// ---- SelfTests/TestCases/TestSuite_Preparation/Helper/PreparationResource.TcPOU
{region 'Documentation'}
(*!
<summary>Controlled local resource for Preparation selftests; only its FB call advances feedback. RequestValue records every command write, including repeated values. Initialize establishes a fresh fixture.</summary>
*)
{endregion}
FUNCTION_BLOCK PreparationResource
VAR_INPUT
    Available : BOOL := TRUE; //! Availability accepted on the next resource-body call.
    Fault : BOOL := FALSE; //! Technical fault accepted on the next resource-body call.
    Advance : BOOL := TRUE; //! FALSE holds feedback without cancelling the accepted request.
END_VAR
VAR
    FActualValue : DINT;
    FRequestedValue : DINT;
    FCommandWriteCount : UDINT;
    FAvailable : BOOL := TRUE;
    FFault : BOOL;
END_VAR

FAvailable := Available;
FFault := Fault;
IF NOT IsReady OR NOT Advance THEN
    RETURN;
END_IF;

IF FActualValue < FRequestedValue THEN
    FActualValue := FActualValue + 1;
ELSIF FActualValue > FRequestedValue THEN
    FActualValue := FActualValue - 1;
END_IF;

{region 'Documentation'}
(*!
<summary>Feedback after the last resource call.</summary>
*)
{endregion}
{attribute 'monitoring' := 'call'}
PROPERTY PUBLIC ActualValue : DINT //! Feedback after the last resource call.
GET // PUBLIC
ActualValue := FActualValue;
END_GET
END_PROPERTY

{region 'Documentation'}
(*!
<summary>Every RequestValue call since fixture initialization, including same-value writes.</summary>
*)
{endregion}
{attribute 'monitoring' := 'call'}
PROPERTY PUBLIC CommandWriteCount : UDINT //! Every RequestValue call since fixture initialization, including same-value writes.
GET // PUBLIC
CommandWriteCount := FCommandWriteCount;
END_GET
END_PROPERTY

{region 'Documentation'}
(*!
<summary>Fault accepted at the last resource call.</summary>
*)
{endregion}
{attribute 'monitoring' := 'call'}
PROPERTY PUBLIC HasError : BOOL //! Fault accepted at the last resource call.
GET // PUBLIC
HasError := FFault;
END_GET
END_PROPERTY

{region 'Documentation'}
(*!
<summary>Restores feedback and request together; fixture setup is not counted as a resource command.</summary>
*)
{endregion}
METHOD PUBLIC Initialize
VAR_INPUT
    InitialValue : DINT; //! Initial feedback and requested target; fixture initialization clears command-write evidence.
END_VAR
FActualValue := InitialValue;
FRequestedValue := InitialValue;
FCommandWriteCount := 0;
FAvailable := TRUE;
FFault := FALSE;
END_METHOD

{region 'Documentation'}
(*!
<summary>Current resource condition permits movement; independent of the target value.</summary>
*)
{endregion}
{attribute 'monitoring' := 'call'}
PROPERTY PUBLIC IsReady : BOOL //! Current resource condition permits movement; independent of the target value.
GET // PUBLIC
IsReady := FAvailable AND NOT FFault;
END_GET
END_PROPERTY

{region 'Documentation'}
(*!
<summary>Last requested target; accepting a command does not establish feedback.</summary>
*)
{endregion}
{attribute 'monitoring' := 'call'}
PROPERTY PUBLIC RequestedValue : DINT //! Last requested target; accepting a command does not establish feedback.
GET // PUBLIC
RequestedValue := FRequestedValue;
END_GET
END_PROPERTY

{region 'Documentation'}
(*!
<summary>Records one command write without changing feedback; a later advancing resource call processes it.</summary>
*)
{endregion}
METHOD PUBLIC RequestValue
VAR_INPUT
    Value : DINT; //! New requested target; this call records a command write without advancing feedback.
END_VAR
FRequestedValue := Value;
FCommandWriteCount := FCommandWriteCount + 1;
END_METHOD

END_FUNCTION_BLOCK

// ---- Framework/Assertions/POU/BasicTypes/DInt/AssertEqual_DInt.TcPOU
{region 'Documentation'}
(*!
<summary>Checks equality with the expected DINT value.</summary>
*)
{endregion}
FUNCTION_BLOCK AssertEqual_DInt EXTENDS AssertionBase
VAR_INPUT
    IN : DINT; //! Actual value checked or observed by this Assertion.
    Expected : DINT; //! Reference value for comparison with IN.
END_VAR

SUPER^();

{region 'Documentation'}
(*!
<summary>Check equality with the expected DINT value.</summary>
*)
{endregion}
METHOD PROTECTED Assert
VAR
    Message : STRING(GVL_Constants.MessageLength);
    ExpectedText : STRING(GVL_Constants.AssertionValueLength);
    ActualText : STRING(GVL_Constants.AssertionValueLength);
END_VAR
IF NOT EvaluationActive THEN
    RETURN;
END_IF;

IF Result = E_Result.Error THEN
    RETURN;
END_IF;

IF Result = E_Result.Failed THEN
    RETURN;
END_IF;

IF IN <> Expected THEN
    ExpectedText := DINT_TO_STRING(Expected);
    ActualText := DINT_TO_STRING(IN);
    Message := CONCAT('Assertion failed: values are not equal. Expected = ',
        ExpectedText);
    Message := CONCAT(Message, ', Actual = ');
    Message := CONCAT(Message, ActualText);
    Message := CONCAT(Message, '.');
    Fail(Message := Message);
    RETURN;
END_IF;

Pass();
END_METHOD

END_FUNCTION_BLOCK

// ---- SelfTests/TestCases/TestSuite_Preparation/Test_PreparationReachesTarget.TcPOU
{region 'Documentation'}
(*!
<summary>Checks real request/feedback separation, multi-cycle target acquisition and already-reached behavior.</summary>
*)
{endregion}
FUNCTION_BLOCK Test_PreparationReachesTarget EXTENDS TestCaseBase
VAR
    FSubject : Prepare_ValueAtTarget;
    FResource : PreparationResource;
    FView : I_Preparation;
    FAlreadyAtTarget : Prepare_ValueAtTarget;
    FObserved : ST_PreparationStatus;
    FExpected : ST_PreparationStatus;
    FObservedEnabled : BOOL;
    FExpectedEnabled : BOOL;
    FCheckPerformed : BOOL;
    FObservedCommandWrites : UDINT;
    FExpectedCommandWrites : UDINT;
    FObservedActualValue : DINT;
    FExpectedActualValue : DINT;
    FObservedRequestedValue : DINT;
    FExpectedRequestedValue : DINT;
    FCheckDiagnosticState : AssertEqual_Int;
    FCheckExecutionStatus : AssertEqual_Int;
    FCheckReady : AssertEqual_Bool;
    FCheckRunning : AssertEqual_Bool;
    FCheckCompleted : AssertEqual_Bool;
    FCheckError : AssertEqual_Bool;
    FCheckEnabled : AssertEqual_Bool;
    FCheckCommandWrites : AssertEqual_UDInt;
    FCheckActualValue : AssertEqual_DInt;
    FCheckRequestedValue : AssertEqual_DInt;
END_VAR
VAR CONSTANT
    CommandAccepted : E_State := E_State.Running;
    ProgressObserved : E_State := E_State.Running + 1;
    TargetReached : E_State := E_State.Running + 2;
    RepeatedCompletion : E_State := E_State.Running + 3;
    AlreadyAtTarget : E_State := E_State.Running + 4;
END_VAR

SUPER^();

{region 'Documentation'}
(*!
<summary>Contributes all owned Assertion results without executing the subjects.</summary>
*)
{endregion}
METHOD PROTECTED AggregateResults
VAR_INPUT
    Aggregator : I_ResultAggregator; //! Borrowed result sink owned by the outer Test Case; add this test's checking Assertions without resetting or retaining the sink.
END_VAR
Aggregator.AddProvider(Provider := FCheckDiagnosticState);
Aggregator.AddProvider(Provider := FCheckExecutionStatus);
Aggregator.AddProvider(Provider := FCheckReady);
Aggregator.AddProvider(Provider := FCheckRunning);
Aggregator.AddProvider(Provider := FCheckCompleted);
Aggregator.AddProvider(Provider := FCheckError);
Aggregator.AddProvider(Provider := FCheckEnabled);
Aggregator.AddProvider(Provider := FCheckCommandWrites);
Aggregator.AddProvider(Provider := FCheckActualValue);
Aggregator.AddProvider(Provider := FCheckRequestedValue);
END_METHOD

{region 'Documentation'}
(*!
<summary>Requires valid base configuration and every owned Assertion.</summary>
*)
{endregion}
METHOD PROTECTED CheckInitialization : BOOL //! TRUE when the inherited initialization check and this concrete fixture check both accept the setup.
CheckInitialization := FALSE;
IF NOT SUPER^.CheckInitialization() THEN
    RETURN;
END_IF;
IF NOT FCheckDiagnosticState.IsInitialized
    OR NOT FCheckExecutionStatus.IsInitialized
    OR NOT FCheckReady.IsInitialized
    OR NOT FCheckRunning.IsInitialized
    OR NOT FCheckCompleted.IsInitialized
    OR NOT FCheckError.IsInitialized
    OR NOT FCheckEnabled.IsInitialized
    OR NOT FCheckCommandWrites.IsInitialized
    OR NOT FCheckActualValue.IsInitialized
    OR NOT FCheckRequestedValue.IsInitialized THEN
    RETURN;
END_IF;

CheckInitialization := TRUE;
END_METHOD

{region 'Documentation'}
(*!
<summary>Configures this scenario, its local subjects and named Assertions.</summary>
*)
{endregion}
METHOD PROTECTED Configure
FPreparationStateCount := 0;
FTestStateCount := 5;
FCheckPerformed := FALSE;
FResource.Initialize(InitialValue := 2);
FSubject.Initialize(Resource := FResource);
FAlreadyAtTarget.Initialize(Resource := FResource);
FView := FSubject;

FCheckDiagnosticState.Initialize(Parent := THIS^,
    AssertionName := 'DiagnosticState');
FCheckExecutionStatus.Initialize(Parent := THIS^,
    AssertionName := 'ExecutionStatus');
FCheckReady.Initialize(Parent := THIS^,
    AssertionName := 'Ready');
FCheckRunning.Initialize(Parent := THIS^,
    AssertionName := 'Running');
FCheckCompleted.Initialize(Parent := THIS^,
    AssertionName := 'Completed');
FCheckError.Initialize(Parent := THIS^,
    AssertionName := 'Error');
FCheckEnabled.Initialize(Parent := THIS^,
    AssertionName := 'Enabled');
FCheckCommandWrites.Initialize(Parent := THIS^,
    AssertionName := 'CommandWrites');
FCheckActualValue.Initialize(Parent := THIS^,
    AssertionName := 'ActualValue');
FCheckRequestedValue.Initialize(Parent := THIS^,
    AssertionName := 'RequestedValue');
END_METHOD

{region 'Documentation'}
(*!
<summary>Ends scenario processing without issuing further resource commands.</summary>
*)
{endregion}
METHOD PROTECTED ProcessAbort
VAR_INPUT
    Enable : BOOL; //! Phase permission supplied by the owning Test Case; FALSE does not authorize progression, while observation may continue.
END_VAR
IF Enable THEN
    CompleteAbort();
END_IF;
END_METHOD

{region 'Documentation'}
(*!
<summary>Compares independent expected values with the captured observations; called when disabled as well.</summary>
*)
{endregion}
METHOD PROTECTED ProcessAssertions
VAR_INPUT
    Enable : BOOL; //! Phase permission supplied by the owning Test Case; FALSE does not authorize progression, while observation may continue.
END_VAR
FCheckDiagnosticState(Enable := Enable,
    State := State,
    IN := TO_INT(FObserved.State),
    Expected := TO_INT(FExpected.State));

FCheckExecutionStatus(Enable := Enable,
    State := State,
    IN := TO_INT(FObserved.ExecutionStatus),
    Expected := TO_INT(FExpected.ExecutionStatus));

FCheckReady(Enable := Enable,
    State := State,
    IN := FObserved.Ready,
    Expected := FExpected.Ready);

FCheckRunning(Enable := Enable,
    State := State,
    IN := FObserved.Running,
    Expected := FExpected.Running);

FCheckCompleted(Enable := Enable,
    State := State,
    IN := FObserved.Completed,
    Expected := FExpected.Completed);

FCheckError(Enable := Enable,
    State := State,
    IN := FObserved.Error,
    Expected := FExpected.Error);

FCheckEnabled(Enable := Enable,
    State := State,
    IN := FObservedEnabled,
    Expected := FExpectedEnabled);

FCheckCommandWrites(Enable := Enable,
    State := State,
    IN := FObservedCommandWrites,
    Expected := FExpectedCommandWrites);

FCheckActualValue(Enable := Enable,
    State := State,
    IN := FObservedActualValue,
    Expected := FExpectedActualValue);

FCheckRequestedValue(Enable := Enable,
    State := State,
    IN := FObservedRequestedValue,
    Expected := FExpectedRequestedValue);

IF Enable
    AND FCheckDiagnosticState.EvaluationActive
    AND FCheckExecutionStatus.EvaluationActive
    AND FCheckReady.EvaluationActive
    AND FCheckRunning.EvaluationActive
    AND FCheckCompleted.EvaluationActive
    AND FCheckError.EvaluationActive
    AND FCheckEnabled.EvaluationActive
    AND FCheckCommandWrites.EvaluationActive
    AND FCheckActualValue.EvaluationActive
    AND FCheckRequestedValue.EvaluationActive THEN
    FCheckPerformed := TRUE;
END_IF;
END_METHOD

{region 'Documentation'}
(*!
<summary>Subjects are exercised by the test, not used as its start prerequisite.</summary>
*)
{endregion}
METHOD PROTECTED ProcessPreparations
VAR_INPUT
    // SA0033: Required hook; this scenario has no Preparation phase.
    {attribute 'analysis' := '-33'}
    Enable : BOOL; //! Phase permission supplied by the owning Test Case; FALSE does not authorize progression, while observation may continue.
END_VAR
END_METHOD

{region 'Documentation'}
(*!
<summary>Restores repeatable fixture state and resets Assertions before returning to Idle.</summary>
*)
{endregion}
METHOD PROTECTED ProcessReset
FCheckPerformed := FALSE;
FResource.Initialize(InitialValue := 2);
FSubject.Initialize(Resource := FResource);
FAlreadyAtTarget.Initialize(Resource := FResource);
FView := FSubject;
FCheckDiagnosticState.Reset();
FCheckExecutionStatus.Reset();
FCheckReady.Reset();
FCheckRunning.Reset();
FCheckCompleted.Reset();
FCheckError.Reset();
FCheckEnabled.Reset();
FCheckCommandWrites.Reset();
FCheckActualValue.Reset();
FCheckRequestedValue.Reset();
CompleteReset();
END_METHOD

{region 'Documentation'}
(*!
<summary>Exercises one named scenario step per call; advances only after actual Assertion evaluation.</summary>
*)
{endregion}
METHOD PROTECTED ProcessTests
VAR_INPUT
    Enable : BOOL; //! Phase permission supplied by the owning Test Case; FALSE does not authorize progression, while observation may continue.
END_VAR
IF NOT Enable THEN
    RETURN;
END_IF;

IF FCheckPerformed THEN
    FCheckPerformed := FALSE;
    IF State = AlreadyAtTarget THEN
        CompleteTests();
        RETURN;
    END_IF;
    NextTestState();
    IF NOT IsTestingActive THEN
        RETURN;
    END_IF;
END_IF;

CASE State OF
    CommandAccepted:
        FResource(Available := TRUE,
            Fault := FALSE,
            Advance := FALSE);
        FSubject(Enable := TRUE,
            TargetValue := 0);
        FExpected.State := E_State.Running;
        FExpected.ExecutionStatus := E_ExecutionStatus.Running;
        FExpected.Ready := FALSE;
        FExpected.Running := TRUE;
        FExpected.Completed := FALSE;
        FExpected.Error := FALSE;
        FExpectedEnabled := TRUE;
        FExpectedCommandWrites := 1;
        FExpectedActualValue := 2;
        FExpectedRequestedValue := 0;

    ProgressObserved:
        FResource(Available := TRUE,
            Fault := FALSE,
            Advance := TRUE);
        FSubject(Enable := TRUE,
            TargetValue := 0);
        FExpected.State := E_State.Running;
        FExpected.ExecutionStatus := E_ExecutionStatus.Running;
        FExpected.Ready := FALSE;
        FExpected.Running := TRUE;
        FExpected.Completed := FALSE;
        FExpected.Error := FALSE;
        FExpectedEnabled := TRUE;
        FExpectedCommandWrites := 1;
        FExpectedActualValue := 1;
        FExpectedRequestedValue := 0;

    TargetReached:
        FResource(Available := TRUE,
            Fault := FALSE,
            Advance := TRUE);
        FSubject(Enable := TRUE,
            TargetValue := 0);
        FExpected.State := E_State.Completed;
        FExpected.ExecutionStatus := E_ExecutionStatus.Completed;
        FExpected.Ready := TRUE;
        FExpected.Running := FALSE;
        FExpected.Completed := TRUE;
        FExpected.Error := FALSE;
        FExpectedEnabled := TRUE;
        FExpectedCommandWrites := 1;
        FExpectedActualValue := 0;
        FExpectedRequestedValue := 0;

    RepeatedCompletion:
        FResource(Available := TRUE,
            Fault := FALSE,
            Advance := TRUE);
        FSubject(Enable := TRUE,
            TargetValue := 0);
        FExpected.State := E_State.Completed;
        FExpected.ExecutionStatus := E_ExecutionStatus.Completed;
        FExpected.Ready := TRUE;
        FExpected.Running := FALSE;
        FExpected.Completed := TRUE;
        FExpected.Error := FALSE;
        FExpectedEnabled := TRUE;
        FExpectedCommandWrites := 1;
        FExpectedActualValue := 0;
        FExpectedRequestedValue := 0;

    AlreadyAtTarget:
        FResource(Available := TRUE,
            Fault := FALSE,
            Advance := TRUE);
        FAlreadyAtTarget(Enable := TRUE,
            TargetValue := 0);
        FView := FAlreadyAtTarget;
        FExpected.State := E_State.Completed;
        FExpected.ExecutionStatus := E_ExecutionStatus.Completed;
        FExpected.Ready := TRUE;
        FExpected.Running := FALSE;
        FExpected.Completed := TRUE;
        FExpected.Error := FALSE;
        FExpectedEnabled := TRUE;
        FExpectedCommandWrites := 1;
        FExpectedActualValue := 0;
        FExpectedRequestedValue := 0;

ELSE
    Error(Message := 'Unexpected Preparation test state.');
    RETURN;
END_CASE;

FObserved := FView.Status;
IF State = AlreadyAtTarget THEN
    FObservedEnabled := FAlreadyAtTarget.Enabled;
ELSE
    FObservedEnabled := FSubject.Enabled;
END_IF;

FObservedCommandWrites := FResource.CommandWriteCount;
FObservedActualValue := FResource.ActualValue;
FObservedRequestedValue := FResource.RequestedValue;
END_METHOD

END_FUNCTION_BLOCK

// ---- SelfTests/TestCases/TestSuite_Preparation/Test_PreparationDisableAndReenable.TcPOU
{region 'Documentation'}
(*!
<summary>Checks that disabling discards local stage progress without cancelling the accepted resource command.</summary>
*)
{endregion}
FUNCTION_BLOCK Test_PreparationDisableAndReenable EXTENDS TestCaseBase
VAR
    FSubject : Prepare_ZeroViaOne;
    FResource : PreparationResource;
    FView : I_Preparation;
    FObserved : ST_PreparationStatus;
    FExpected : ST_PreparationStatus;
    FObservedEnabled : BOOL;
    FExpectedEnabled : BOOL;
    FCheckPerformed : BOOL;
    FObservedCommandWrites : UDINT;
    FExpectedCommandWrites : UDINT;
    FObservedActualValue : DINT;
    FExpectedActualValue : DINT;
    FObservedRequestedValue : DINT;
    FExpectedRequestedValue : DINT;
    FCheckDiagnosticState : AssertEqual_Int;
    FCheckExecutionStatus : AssertEqual_Int;
    FCheckReady : AssertEqual_Bool;
    FCheckRunning : AssertEqual_Bool;
    FCheckCompleted : AssertEqual_Bool;
    FCheckError : AssertEqual_Bool;
    FCheckEnabled : AssertEqual_Bool;
    FCheckCommandWrites : AssertEqual_UDInt;
    FCheckActualValue : AssertEqual_DInt;
    FCheckRequestedValue : AssertEqual_DInt;
END_VAR
VAR CONSTANT
    IntermediateRequested : E_State := E_State.Running;
    DisableDuringMovement : E_State := E_State.Running + 1;
    AcceptedRequestContinues : E_State := E_State.Running + 2;
    ResourceChangedWhileDisabled : E_State := E_State.Running + 3;
    ReenableFromCurrentFeedback : E_State := E_State.Running + 4;
    IntermediateApproached : E_State := E_State.Running + 5;
    FinalTargetRequested : E_State := E_State.Running + 6;
    FinalTargetReached : E_State := E_State.Running + 7;
END_VAR

SUPER^();

{region 'Documentation'}
(*!
<summary>Contributes all owned Assertion results without executing the subjects.</summary>
*)
{endregion}
METHOD PROTECTED AggregateResults
VAR_INPUT
    Aggregator : I_ResultAggregator; //! Borrowed result sink owned by the outer Test Case; add this test's checking Assertions without resetting or retaining the sink.
END_VAR
Aggregator.AddProvider(Provider := FCheckDiagnosticState);
Aggregator.AddProvider(Provider := FCheckExecutionStatus);
Aggregator.AddProvider(Provider := FCheckReady);
Aggregator.AddProvider(Provider := FCheckRunning);
Aggregator.AddProvider(Provider := FCheckCompleted);
Aggregator.AddProvider(Provider := FCheckError);
Aggregator.AddProvider(Provider := FCheckEnabled);
Aggregator.AddProvider(Provider := FCheckCommandWrites);
Aggregator.AddProvider(Provider := FCheckActualValue);
Aggregator.AddProvider(Provider := FCheckRequestedValue);
END_METHOD

{region 'Documentation'}
(*!
<summary>Requires valid base configuration and every owned Assertion.</summary>
*)
{endregion}
METHOD PROTECTED CheckInitialization : BOOL //! TRUE when the inherited initialization check and this concrete fixture check both accept the setup.
CheckInitialization := FALSE;
IF NOT SUPER^.CheckInitialization() THEN
    RETURN;
END_IF;
IF NOT FCheckDiagnosticState.IsInitialized
    OR NOT FCheckExecutionStatus.IsInitialized
    OR NOT FCheckReady.IsInitialized
    OR NOT FCheckRunning.IsInitialized
    OR NOT FCheckCompleted.IsInitialized
    OR NOT FCheckError.IsInitialized
    OR NOT FCheckEnabled.IsInitialized
    OR NOT FCheckCommandWrites.IsInitialized
    OR NOT FCheckActualValue.IsInitialized
    OR NOT FCheckRequestedValue.IsInitialized THEN
    RETURN;
END_IF;

CheckInitialization := TRUE;
END_METHOD

{region 'Documentation'}
(*!
<summary>Configures this scenario, its local subjects and named Assertions.</summary>
*)
{endregion}
METHOD PROTECTED Configure
FPreparationStateCount := 0;
FTestStateCount := 8;
FCheckPerformed := FALSE;
FResource.Initialize(InitialValue := 3);
FSubject.Initialize(Resource := FResource);
FView := FSubject;

FCheckDiagnosticState.Initialize(Parent := THIS^,
    AssertionName := 'DiagnosticState');
FCheckExecutionStatus.Initialize(Parent := THIS^,
    AssertionName := 'ExecutionStatus');
FCheckReady.Initialize(Parent := THIS^,
    AssertionName := 'Ready');
FCheckRunning.Initialize(Parent := THIS^,
    AssertionName := 'Running');
FCheckCompleted.Initialize(Parent := THIS^,
    AssertionName := 'Completed');
FCheckError.Initialize(Parent := THIS^,
    AssertionName := 'Error');
FCheckEnabled.Initialize(Parent := THIS^,
    AssertionName := 'Enabled');
FCheckCommandWrites.Initialize(Parent := THIS^,
    AssertionName := 'CommandWrites');
FCheckActualValue.Initialize(Parent := THIS^,
    AssertionName := 'ActualValue');
FCheckRequestedValue.Initialize(Parent := THIS^,
    AssertionName := 'RequestedValue');
END_METHOD

{region 'Documentation'}
(*!
<summary>Ends scenario processing without issuing further resource commands.</summary>
*)
{endregion}
METHOD PROTECTED ProcessAbort
VAR_INPUT
    Enable : BOOL; //! Phase permission supplied by the owning Test Case; FALSE does not authorize progression, while observation may continue.
END_VAR
IF Enable THEN
    CompleteAbort();
END_IF;
END_METHOD

{region 'Documentation'}
(*!
<summary>Compares independent expected values with the captured observations; called when disabled as well.</summary>
*)
{endregion}
METHOD PROTECTED ProcessAssertions
VAR_INPUT
    Enable : BOOL; //! Phase permission supplied by the owning Test Case; FALSE does not authorize progression, while observation may continue.
END_VAR
FCheckDiagnosticState(Enable := Enable,
    State := State,
    IN := TO_INT(FObserved.State),
    Expected := TO_INT(FExpected.State));

FCheckExecutionStatus(Enable := Enable,
    State := State,
    IN := TO_INT(FObserved.ExecutionStatus),
    Expected := TO_INT(FExpected.ExecutionStatus));

FCheckReady(Enable := Enable,
    State := State,
    IN := FObserved.Ready,
    Expected := FExpected.Ready);

FCheckRunning(Enable := Enable,
    State := State,
    IN := FObserved.Running,
    Expected := FExpected.Running);

FCheckCompleted(Enable := Enable,
    State := State,
    IN := FObserved.Completed,
    Expected := FExpected.Completed);

FCheckError(Enable := Enable,
    State := State,
    IN := FObserved.Error,
    Expected := FExpected.Error);

FCheckEnabled(Enable := Enable,
    State := State,
    IN := FObservedEnabled,
    Expected := FExpectedEnabled);

FCheckCommandWrites(Enable := Enable,
    State := State,
    IN := FObservedCommandWrites,
    Expected := FExpectedCommandWrites);

FCheckActualValue(Enable := Enable,
    State := State,
    IN := FObservedActualValue,
    Expected := FExpectedActualValue);

FCheckRequestedValue(Enable := Enable,
    State := State,
    IN := FObservedRequestedValue,
    Expected := FExpectedRequestedValue);

IF Enable
    AND FCheckDiagnosticState.EvaluationActive
    AND FCheckExecutionStatus.EvaluationActive
    AND FCheckReady.EvaluationActive
    AND FCheckRunning.EvaluationActive
    AND FCheckCompleted.EvaluationActive
    AND FCheckError.EvaluationActive
    AND FCheckEnabled.EvaluationActive
    AND FCheckCommandWrites.EvaluationActive
    AND FCheckActualValue.EvaluationActive
    AND FCheckRequestedValue.EvaluationActive THEN
    FCheckPerformed := TRUE;
END_IF;
END_METHOD

{region 'Documentation'}
(*!
<summary>Subjects are exercised by the test, not used as its start prerequisite.</summary>
*)
{endregion}
METHOD PROTECTED ProcessPreparations
VAR_INPUT
    // SA0033: Required hook; this scenario has no Preparation phase.
    {attribute 'analysis' := '-33'}
    Enable : BOOL; //! Phase permission supplied by the owning Test Case; FALSE does not authorize progression, while observation may continue.
END_VAR
END_METHOD

{region 'Documentation'}
(*!
<summary>Restores repeatable fixture state and resets Assertions before returning to Idle.</summary>
*)
{endregion}
METHOD PROTECTED ProcessReset
FCheckPerformed := FALSE;
FResource.Initialize(InitialValue := 3);
FSubject.Initialize(Resource := FResource);
FView := FSubject;
FCheckDiagnosticState.Reset();
FCheckExecutionStatus.Reset();
FCheckReady.Reset();
FCheckRunning.Reset();
FCheckCompleted.Reset();
FCheckError.Reset();
FCheckEnabled.Reset();
FCheckCommandWrites.Reset();
FCheckActualValue.Reset();
FCheckRequestedValue.Reset();
CompleteReset();
END_METHOD

{region 'Documentation'}
(*!
<summary>Exercises one named scenario step per call; advances only after actual Assertion evaluation.</summary>
*)
{endregion}
METHOD PROTECTED ProcessTests
VAR_INPUT
    Enable : BOOL; //! Phase permission supplied by the owning Test Case; FALSE does not authorize progression, while observation may continue.
END_VAR
IF NOT Enable THEN
    RETURN;
END_IF;

IF FCheckPerformed THEN
    FCheckPerformed := FALSE;
    IF State = FinalTargetReached THEN
        CompleteTests();
        RETURN;
    END_IF;
    NextTestState();
    IF NOT IsTestingActive THEN
        RETURN;
    END_IF;
END_IF;

CASE State OF
    IntermediateRequested:
        FResource(Available := TRUE,
            Fault := FALSE,
            Advance := FALSE);
        FSubject(Enable := TRUE);
        FExpected.State := E_State.Preparing;
        FExpected.ExecutionStatus := E_ExecutionStatus.Running;
        FExpected.Ready := FALSE;
        FExpected.Running := TRUE;
        FExpected.Completed := FALSE;
        FExpected.Error := FALSE;
        FExpectedEnabled := TRUE;
        FExpectedCommandWrites := 1;
        FExpectedActualValue := 3;
        FExpectedRequestedValue := 1;

    DisableDuringMovement:
        FResource(Available := TRUE,
            Fault := FALSE,
            Advance := TRUE);
        FSubject(Enable := FALSE);
        FExpected.State := E_State.Idle;
        FExpected.ExecutionStatus := E_ExecutionStatus.Idle;
        FExpected.Ready := TRUE;
        FExpected.Running := FALSE;
        FExpected.Completed := FALSE;
        FExpected.Error := FALSE;
        FExpectedEnabled := FALSE;
        FExpectedCommandWrites := 1;
        FExpectedActualValue := 2;
        FExpectedRequestedValue := 1;

    AcceptedRequestContinues:
        FResource(Available := TRUE,
            Fault := FALSE,
            Advance := TRUE);
        FSubject(Enable := FALSE);
        FExpected.State := E_State.Idle;
        FExpected.ExecutionStatus := E_ExecutionStatus.Idle;
        FExpected.Ready := TRUE;
        FExpected.Running := FALSE;
        FExpected.Completed := FALSE;
        FExpected.Error := FALSE;
        FExpectedEnabled := FALSE;
        FExpectedCommandWrites := 1;
        FExpectedActualValue := 1;
        FExpectedRequestedValue := 1;

    ResourceChangedWhileDisabled:
        FResource.RequestValue(Value := 3);
        FResource(Available := TRUE,
            Fault := FALSE,
            Advance := TRUE);
        FSubject(Enable := FALSE);
        FExpected.State := E_State.Idle;
        FExpected.ExecutionStatus := E_ExecutionStatus.Idle;
        FExpected.Ready := TRUE;
        FExpected.Running := FALSE;
        FExpected.Completed := FALSE;
        FExpected.Error := FALSE;
        FExpectedEnabled := FALSE;
        FExpectedCommandWrites := 2;
        FExpectedActualValue := 2;
        FExpectedRequestedValue := 3;

    ReenableFromCurrentFeedback:
        FResource(Available := TRUE,
            Fault := FALSE,
            Advance := TRUE);
        FSubject(Enable := TRUE);
        FExpected.State := E_State.Preparing;
        FExpected.ExecutionStatus := E_ExecutionStatus.Running;
        FExpected.Ready := FALSE;
        FExpected.Running := TRUE;
        FExpected.Completed := FALSE;
        FExpected.Error := FALSE;
        FExpectedEnabled := TRUE;
        FExpectedCommandWrites := 3;
        FExpectedActualValue := 3;
        FExpectedRequestedValue := 1;

    IntermediateApproached:
        FResource(Available := TRUE,
            Fault := FALSE,
            Advance := TRUE);
        FSubject(Enable := TRUE);
        FExpected.State := E_State.Preparing;
        FExpected.ExecutionStatus := E_ExecutionStatus.Running;
        FExpected.Ready := FALSE;
        FExpected.Running := TRUE;
        FExpected.Completed := FALSE;
        FExpected.Error := FALSE;
        FExpectedEnabled := TRUE;
        FExpectedCommandWrites := 3;
        FExpectedActualValue := 2;
        FExpectedRequestedValue := 1;

    FinalTargetRequested:
        FResource(Available := TRUE,
            Fault := FALSE,
            Advance := TRUE);
        FSubject(Enable := TRUE);
        FExpected.State := E_State.Running;
        FExpected.ExecutionStatus := E_ExecutionStatus.Running;
        FExpected.Ready := FALSE;
        FExpected.Running := TRUE;
        FExpected.Completed := FALSE;
        FExpected.Error := FALSE;
        FExpectedEnabled := TRUE;
        FExpectedCommandWrites := 4;
        FExpectedActualValue := 1;
        FExpectedRequestedValue := 0;

    FinalTargetReached:
        FResource(Available := TRUE,
            Fault := FALSE,
            Advance := TRUE);
        FSubject(Enable := TRUE);
        FExpected.State := E_State.Completed;
        FExpected.ExecutionStatus := E_ExecutionStatus.Completed;
        FExpected.Ready := TRUE;
        FExpected.Running := FALSE;
        FExpected.Completed := TRUE;
        FExpected.Error := FALSE;
        FExpectedEnabled := TRUE;
        FExpectedCommandWrites := 4;
        FExpectedActualValue := 0;
        FExpectedRequestedValue := 0;

ELSE
    Error(Message := 'Unexpected Preparation test state.');
    RETURN;
END_CASE;

FObserved := FView.Status;
FObservedEnabled := FSubject.Enabled;

FObservedCommandWrites := FResource.CommandWriteCount;
FObservedActualValue := FResource.ActualValue;
FObservedRequestedValue := FResource.RequestedValue;
END_METHOD

END_FUNCTION_BLOCK

// ---- SelfTests/TestCases/TestSuite_Preparation/Helper/Prepare_ZeroViaOne.TcPOU
{region 'Documentation'}
(*!
<summary>Stateful local Preparation: establish value one before commanding zero. Disabled calls discard local progress without cancelling the resource request.</summary>
*)
{endregion}
FUNCTION_BLOCK Prepare_ZeroViaOne EXTENDS PreparationBase
VAR
    FResource : REFERENCE TO PreparationResource;
    FProgress : E_State := E_State.Idle;
END_VAR

VAR CONSTANT
    IntermediateValue : DINT := 1;
    TargetValue : DINT := 0;
END_VAR

SUPER^();

{region 'Documentation'}
(*!
<summary>Binds a static test-owned resource and clears local sequence progress.</summary>
*)
{endregion}
METHOD PUBLIC Initialize
VAR_IN_OUT
    // SA0167: Borrowed static resource, not a temporary instance.
    {attribute 'analysis' := '-167'}
    Resource : PreparationResource; //! Borrowed static resource retained by reference; keep it alive and stable for all preparation calls.
END_VAR
FResource REF= Resource;
FProgress := E_State.Idle;
END_METHOD

{region 'Documentation'}
(*!
<summary>Observes current feedback; enabling permits the two-stage resource sequence.</summary>
*)
{endregion}
METHOD PROTECTED Prepare
IF NOT Enabled THEN
    FProgress := E_State.Idle;
END_IF;
IF NOT __ISVALIDREF(FResource) THEN
    UpdateStatus(State := E_State.Error,
        ExecutionStatus := E_ExecutionStatus.Error,
        Ready := FALSE);
    RETURN;
END_IF;
IF FResource.HasError THEN
    UpdateStatus(State := E_State.Error,
        ExecutionStatus := E_ExecutionStatus.Error,
        Ready := FALSE);
    RETURN;
END_IF;

IF (FResource.ActualValue = TargetValue) AND (FResource.RequestedValue = TargetValue) THEN
    UpdateStatus(State := E_State.Completed,
        ExecutionStatus := E_ExecutionStatus.Completed,
        Ready := FResource.IsReady);
ELSIF Enabled AND FResource.IsReady THEN
    StateMachine();
    IF FProgress = E_State.Error THEN
        UpdateStatus(State := E_State.Error,
            ExecutionStatus := E_ExecutionStatus.Error,
            Ready := FALSE);
    ELSE
        UpdateStatus(State := FProgress,
            ExecutionStatus := E_ExecutionStatus.Running,
            Ready := FALSE);
    END_IF;
ELSIF FResource.IsReady THEN
    UpdateStatus(State := E_State.Idle,
        ExecutionStatus := E_ExecutionStatus.Idle,
        Ready := TRUE);
ELSE
    UpdateStatus(State := E_State.Idle,
        ExecutionStatus := E_ExecutionStatus.NotReady,
        Ready := FALSE);
END_IF;
END_METHOD

{region 'Documentation'}
(*!
<summary>Advances at most one resource stage per call; no feedback simulation.</summary>
*)
{endregion}
METHOD PRIVATE StateMachine
CASE FProgress OF
    E_State.Idle:
        IF FResource.ActualValue = IntermediateValue THEN
            FResource.RequestValue(Value := TargetValue);
            FProgress := E_State.Running;
        ELSE
            FResource.RequestValue(Value := IntermediateValue);
            FProgress := E_State.Preparing;
        END_IF;

    E_State.Preparing:
        IF FResource.ActualValue = IntermediateValue THEN
            FResource.RequestValue(Value := TargetValue);
            FProgress := E_State.Running;
        END_IF;

    E_State.Running:
        RETURN;
ELSE
    FProgress := E_State.Error;
END_CASE;
END_METHOD

END_FUNCTION_BLOCK

// ---- SelfTests/TestCases/TestSuite_Preparation/Test_PreparationCompletionTracksTarget.TcPOU
{region 'Documentation'}
(*!
<summary>Checks real Preparation-to-test handover; loss of Ready/Completed does not restart or block the active Test Case.</summary>
*)
{endregion}
FUNCTION_BLOCK Test_PreparationCompletionTracksTarget EXTENDS TestCaseBase
VAR
    FSubject : Prepare_ValueAtTarget;
    FResource : PreparationResource;
    FView : I_Preparation;
    FResourceAvailable : BOOL := TRUE;
    FObserved : ST_PreparationStatus;
    FExpected : ST_PreparationStatus;
    FObservedEnabled : BOOL;
    FExpectedEnabled : BOOL;
    FCheckPerformed : BOOL;
    FObservedCommandWrites : UDINT;
    FExpectedCommandWrites : UDINT;
    FObservedActualValue : DINT;
    FExpectedActualValue : DINT;
    FObservedRequestedValue : DINT;
    FExpectedRequestedValue : DINT;
    FCheckDiagnosticState : AssertEqual_Int;
    FCheckExecutionStatus : AssertEqual_Int;
    FCheckReady : AssertEqual_Bool;
    FCheckRunning : AssertEqual_Bool;
    FCheckCompleted : AssertEqual_Bool;
    FCheckError : AssertEqual_Bool;
    FCheckEnabled : AssertEqual_Bool;
    FCheckCommandWrites : AssertEqual_UDInt;
    FCheckActualValue : AssertEqual_DInt;
    FCheckRequestedValue : AssertEqual_DInt;
    FCheckTestingActive : AssertEqual_Bool;
END_VAR
VAR CONSTANT
    PreparationHandedOver : E_State := E_State.Running;
    TargetAndReadinessLost : E_State := E_State.Running + 1;
    TestingContinues : E_State := E_State.Running + 2;
END_VAR

SUPER^();

{region 'Documentation'}
(*!
<summary>Contributes all owned Assertion results without executing the subjects.</summary>
*)
{endregion}
METHOD PROTECTED AggregateResults
VAR_INPUT
    Aggregator : I_ResultAggregator; //! Borrowed result sink owned by the outer Test Case; add this test's checking Assertions without resetting or retaining the sink.
END_VAR
Aggregator.AddProvider(Provider := FCheckDiagnosticState);
Aggregator.AddProvider(Provider := FCheckExecutionStatus);
Aggregator.AddProvider(Provider := FCheckReady);
Aggregator.AddProvider(Provider := FCheckRunning);
Aggregator.AddProvider(Provider := FCheckCompleted);
Aggregator.AddProvider(Provider := FCheckError);
Aggregator.AddProvider(Provider := FCheckEnabled);
Aggregator.AddProvider(Provider := FCheckCommandWrites);
Aggregator.AddProvider(Provider := FCheckActualValue);
Aggregator.AddProvider(Provider := FCheckRequestedValue);
Aggregator.AddProvider(Provider := FCheckTestingActive);
END_METHOD

{region 'Documentation'}
(*!
<summary>Requires valid base configuration and every owned Assertion.</summary>
*)
{endregion}
METHOD PROTECTED CheckInitialization : BOOL //! TRUE when the inherited initialization check and this concrete fixture check both accept the setup.
CheckInitialization := FALSE;
IF NOT SUPER^.CheckInitialization() THEN
    RETURN;
END_IF;
IF NOT FCheckDiagnosticState.IsInitialized
    OR NOT FCheckExecutionStatus.IsInitialized
    OR NOT FCheckReady.IsInitialized
    OR NOT FCheckRunning.IsInitialized
    OR NOT FCheckCompleted.IsInitialized
    OR NOT FCheckError.IsInitialized
    OR NOT FCheckEnabled.IsInitialized
    OR NOT FCheckCommandWrites.IsInitialized
    OR NOT FCheckActualValue.IsInitialized
    OR NOT FCheckRequestedValue.IsInitialized
    OR NOT FCheckTestingActive.IsInitialized THEN
    RETURN;
END_IF;

CheckInitialization := TRUE;
END_METHOD

{region 'Documentation'}
(*!
<summary>Configures this scenario, its local subjects and named Assertions.</summary>
*)
{endregion}
METHOD PROTECTED Configure
FPreparationStateCount := 1;
FTestStateCount := 3;
FCheckPerformed := FALSE;
FResource.Initialize(InitialValue := 2);
FSubject.Initialize(Resource := FResource);
FView := FSubject;
FResourceAvailable := TRUE;

FCheckDiagnosticState.Initialize(Parent := THIS^,
    AssertionName := 'DiagnosticState');
FCheckExecutionStatus.Initialize(Parent := THIS^,
    AssertionName := 'ExecutionStatus');
FCheckReady.Initialize(Parent := THIS^,
    AssertionName := 'Ready');
FCheckRunning.Initialize(Parent := THIS^,
    AssertionName := 'Running');
FCheckCompleted.Initialize(Parent := THIS^,
    AssertionName := 'Completed');
FCheckError.Initialize(Parent := THIS^,
    AssertionName := 'Error');
FCheckEnabled.Initialize(Parent := THIS^,
    AssertionName := 'Enabled');
FCheckCommandWrites.Initialize(Parent := THIS^,
    AssertionName := 'CommandWrites');
FCheckActualValue.Initialize(Parent := THIS^,
    AssertionName := 'ActualValue');
FCheckRequestedValue.Initialize(Parent := THIS^,
    AssertionName := 'RequestedValue');
FCheckTestingActive.Initialize(Parent := THIS^,
    AssertionName := 'TestingActive');
END_METHOD

{region 'Documentation'}
(*!
<summary>Ends scenario processing without issuing further resource commands.</summary>
*)
{endregion}
METHOD PROTECTED ProcessAbort
VAR_INPUT
    Enable : BOOL; //! Phase permission supplied by the owning Test Case; FALSE does not authorize progression, while observation may continue.
END_VAR
IF Enable THEN
    CompleteAbort();
END_IF;
END_METHOD

{region 'Documentation'}
(*!
<summary>Compares independent expected values with the captured observations; called when disabled as well.</summary>
*)
{endregion}
METHOD PROTECTED ProcessAssertions
VAR_INPUT
    Enable : BOOL; //! Phase permission supplied by the owning Test Case; FALSE does not authorize progression, while observation may continue.
END_VAR
FCheckDiagnosticState(Enable := Enable,
    State := State,
    IN := TO_INT(FObserved.State),
    Expected := TO_INT(FExpected.State));

FCheckExecutionStatus(Enable := Enable,
    State := State,
    IN := TO_INT(FObserved.ExecutionStatus),
    Expected := TO_INT(FExpected.ExecutionStatus));

FCheckReady(Enable := Enable,
    State := State,
    IN := FObserved.Ready,
    Expected := FExpected.Ready);

FCheckRunning(Enable := Enable,
    State := State,
    IN := FObserved.Running,
    Expected := FExpected.Running);

FCheckCompleted(Enable := Enable,
    State := State,
    IN := FObserved.Completed,
    Expected := FExpected.Completed);

FCheckError(Enable := Enable,
    State := State,
    IN := FObserved.Error,
    Expected := FExpected.Error);

FCheckEnabled(Enable := Enable,
    State := State,
    IN := FObservedEnabled,
    Expected := FExpectedEnabled);

FCheckCommandWrites(Enable := Enable,
    State := State,
    IN := FObservedCommandWrites,
    Expected := FExpectedCommandWrites);

FCheckActualValue(Enable := Enable,
    State := State,
    IN := FObservedActualValue,
    Expected := FExpectedActualValue);

FCheckRequestedValue(Enable := Enable,
    State := State,
    IN := FObservedRequestedValue,
    Expected := FExpectedRequestedValue);

FCheckTestingActive(Enable := Enable,
    State := State,
    IN := IsTestingActive,
    Expected := TRUE);

IF Enable
    AND FCheckDiagnosticState.EvaluationActive
    AND FCheckExecutionStatus.EvaluationActive
    AND FCheckReady.EvaluationActive
    AND FCheckRunning.EvaluationActive
    AND FCheckCompleted.EvaluationActive
    AND FCheckError.EvaluationActive
    AND FCheckEnabled.EvaluationActive
    AND FCheckCommandWrites.EvaluationActive
    AND FCheckActualValue.EvaluationActive
    AND FCheckRequestedValue.EvaluationActive
    AND FCheckTestingActive.EvaluationActive THEN
    FCheckPerformed := TRUE;
END_IF;
END_METHOD

{region 'Documentation'}
(*!
<summary>Runs the real Preparation phase and projects its observations to the owner.</summary>
*)
{endregion}
METHOD PROTECTED ProcessPreparations
VAR_INPUT
    Enable : BOOL; //! Phase permission supplied by the owning Test Case; FALSE does not authorize progression, while observation may continue.
END_VAR
FResource(Available := FResourceAvailable,
    Fault := FALSE,
    Advance := TRUE);
FSubject(Enable := Enable,
    TargetValue := 0);
FObserved := FView.Status;
UpdatePreparationStatus(Ready := FObserved.Ready,
    Running := FObserved.Running,
    Completed := FObserved.Completed,
    HasError := FObserved.Error,
    State := FObserved.State);
END_METHOD

{region 'Documentation'}
(*!
<summary>Restores repeatable fixture state and resets Assertions before returning to Idle.</summary>
*)
{endregion}
METHOD PROTECTED ProcessReset
FCheckPerformed := FALSE;
FResource.Initialize(InitialValue := 2);
FSubject.Initialize(Resource := FResource);
FView := FSubject;
FResourceAvailable := TRUE;
FCheckDiagnosticState.Reset();
FCheckExecutionStatus.Reset();
FCheckReady.Reset();
FCheckRunning.Reset();
FCheckCompleted.Reset();
FCheckError.Reset();
FCheckEnabled.Reset();
FCheckCommandWrites.Reset();
FCheckActualValue.Reset();
FCheckRequestedValue.Reset();
FCheckTestingActive.Reset();
CompleteReset();
END_METHOD

{region 'Documentation'}
(*!
<summary>Exercises one named scenario step per call; advances only after actual Assertion evaluation.</summary>
*)
{endregion}
METHOD PROTECTED ProcessTests
VAR_INPUT
    Enable : BOOL; //! Phase permission supplied by the owning Test Case; FALSE does not authorize progression, while observation may continue.
END_VAR
IF NOT Enable THEN
    RETURN;
END_IF;

IF FCheckPerformed THEN
    FCheckPerformed := FALSE;
    IF State = TestingContinues THEN
        CompleteTests();
        RETURN;
    END_IF;
    NextTestState();
    IF NOT IsTestingActive THEN
        RETURN;
    END_IF;
END_IF;

CASE State OF
    PreparationHandedOver:
        FResource.RequestValue(Value := 2);
        FResourceAvailable := FALSE;
        FExpected.State := E_State.Completed;
        FExpected.ExecutionStatus := E_ExecutionStatus.Completed;
        FExpected.Ready := TRUE;
        FExpected.Running := FALSE;
        FExpected.Completed := TRUE;
        FExpected.Error := FALSE;
        FExpectedEnabled := FALSE;
        FExpectedCommandWrites := 2;
        FExpectedActualValue := 0;
        FExpectedRequestedValue := 2;

    TargetAndReadinessLost:
        FExpected.State := E_State.Idle;
        FExpected.ExecutionStatus := E_ExecutionStatus.NotReady;
        FExpected.Ready := FALSE;
        FExpected.Running := FALSE;
        FExpected.Completed := FALSE;
        FExpected.Error := FALSE;
        FExpectedEnabled := FALSE;
        FExpectedCommandWrites := 2;
        FExpectedActualValue := 0;
        FExpectedRequestedValue := 2;

    TestingContinues:
        FExpected.State := E_State.Idle;
        FExpected.ExecutionStatus := E_ExecutionStatus.NotReady;
        FExpected.Ready := FALSE;
        FExpected.Running := FALSE;
        FExpected.Completed := FALSE;
        FExpected.Error := FALSE;
        FExpectedEnabled := FALSE;
        FExpectedCommandWrites := 2;
        FExpectedActualValue := 0;
        FExpectedRequestedValue := 2;

ELSE
    Error(Message := 'Unexpected Preparation test state.');
    RETURN;
END_CASE;

FObserved := FView.Status;
FObservedEnabled := FSubject.Enabled;

FObservedCommandWrites := FResource.CommandWriteCount;
FObservedActualValue := FResource.ActualValue;
FObservedRequestedValue := FResource.RequestedValue;
END_METHOD

END_FUNCTION_BLOCK

// ---- SelfTests/TestCases/TestSuite_Preparation/Test_PreparationResourceError.TcPOU
{region 'Documentation'}
(*!
<summary>Checks resource faults before actions, during progress and after completion, without failing the outer Test Case.</summary>
*)
{endregion}
FUNCTION_BLOCK Test_PreparationResourceError EXTENDS TestCaseBase
VAR
    FSubject : Prepare_ValueAtTarget;
    FResource : PreparationResource;
    FView : I_Preparation;
    FObserved : ST_PreparationStatus;
    FExpected : ST_PreparationStatus;
    FObservedEnabled : BOOL;
    FExpectedEnabled : BOOL;
    FCheckPerformed : BOOL;
    FObservedCommandWrites : UDINT;
    FExpectedCommandWrites : UDINT;
    FObservedActualValue : DINT;
    FExpectedActualValue : DINT;
    FObservedRequestedValue : DINT;
    FExpectedRequestedValue : DINT;
    FCheckDiagnosticState : AssertEqual_Int;
    FCheckExecutionStatus : AssertEqual_Int;
    FCheckReady : AssertEqual_Bool;
    FCheckRunning : AssertEqual_Bool;
    FCheckCompleted : AssertEqual_Bool;
    FCheckError : AssertEqual_Bool;
    FCheckEnabled : AssertEqual_Bool;
    FCheckCommandWrites : AssertEqual_UDInt;
    FCheckActualValue : AssertEqual_DInt;
    FCheckRequestedValue : AssertEqual_DInt;
END_VAR
VAR CONSTANT
    FaultBeforeAction : E_State := E_State.Running;
    RecoveredRequest : E_State := E_State.Running + 1;
    FaultDuringProgress : E_State := E_State.Running + 2;
    RecoveredProgress : E_State := E_State.Running + 3;
    RecoveredTarget : E_State := E_State.Running + 4;
    FaultAfterCompletion : E_State := E_State.Running + 5;
    CompletionWithoutReadiness : E_State := E_State.Running + 6;
END_VAR

SUPER^();

{region 'Documentation'}
(*!
<summary>Contributes all owned Assertion results without executing the subjects.</summary>
*)
{endregion}
METHOD PROTECTED AggregateResults
VAR_INPUT
    Aggregator : I_ResultAggregator; //! Borrowed result sink owned by the outer Test Case; add this test's checking Assertions without resetting or retaining the sink.
END_VAR
Aggregator.AddProvider(Provider := FCheckDiagnosticState);
Aggregator.AddProvider(Provider := FCheckExecutionStatus);
Aggregator.AddProvider(Provider := FCheckReady);
Aggregator.AddProvider(Provider := FCheckRunning);
Aggregator.AddProvider(Provider := FCheckCompleted);
Aggregator.AddProvider(Provider := FCheckError);
Aggregator.AddProvider(Provider := FCheckEnabled);
Aggregator.AddProvider(Provider := FCheckCommandWrites);
Aggregator.AddProvider(Provider := FCheckActualValue);
Aggregator.AddProvider(Provider := FCheckRequestedValue);
END_METHOD

{region 'Documentation'}
(*!
<summary>Requires valid base configuration and every owned Assertion.</summary>
*)
{endregion}
METHOD PROTECTED CheckInitialization : BOOL //! TRUE when the inherited initialization check and this concrete fixture check both accept the setup.
CheckInitialization := FALSE;
IF NOT SUPER^.CheckInitialization() THEN
    RETURN;
END_IF;
IF NOT FCheckDiagnosticState.IsInitialized
    OR NOT FCheckExecutionStatus.IsInitialized
    OR NOT FCheckReady.IsInitialized
    OR NOT FCheckRunning.IsInitialized
    OR NOT FCheckCompleted.IsInitialized
    OR NOT FCheckError.IsInitialized
    OR NOT FCheckEnabled.IsInitialized
    OR NOT FCheckCommandWrites.IsInitialized
    OR NOT FCheckActualValue.IsInitialized
    OR NOT FCheckRequestedValue.IsInitialized THEN
    RETURN;
END_IF;

CheckInitialization := TRUE;
END_METHOD

{region 'Documentation'}
(*!
<summary>Configures this scenario, its local subjects and named Assertions.</summary>
*)
{endregion}
METHOD PROTECTED Configure
FPreparationStateCount := 0;
FTestStateCount := 7;
FCheckPerformed := FALSE;
FResource.Initialize(InitialValue := 2);
FSubject.Initialize(Resource := FResource);
FView := FSubject;

FCheckDiagnosticState.Initialize(Parent := THIS^,
    AssertionName := 'DiagnosticState');
FCheckExecutionStatus.Initialize(Parent := THIS^,
    AssertionName := 'ExecutionStatus');
FCheckReady.Initialize(Parent := THIS^,
    AssertionName := 'Ready');
FCheckRunning.Initialize(Parent := THIS^,
    AssertionName := 'Running');
FCheckCompleted.Initialize(Parent := THIS^,
    AssertionName := 'Completed');
FCheckError.Initialize(Parent := THIS^,
    AssertionName := 'Error');
FCheckEnabled.Initialize(Parent := THIS^,
    AssertionName := 'Enabled');
FCheckCommandWrites.Initialize(Parent := THIS^,
    AssertionName := 'CommandWrites');
FCheckActualValue.Initialize(Parent := THIS^,
    AssertionName := 'ActualValue');
FCheckRequestedValue.Initialize(Parent := THIS^,
    AssertionName := 'RequestedValue');
END_METHOD

{region 'Documentation'}
(*!
<summary>Ends scenario processing without issuing further resource commands.</summary>
*)
{endregion}
METHOD PROTECTED ProcessAbort
VAR_INPUT
    Enable : BOOL; //! Phase permission supplied by the owning Test Case; FALSE does not authorize progression, while observation may continue.
END_VAR
IF Enable THEN
    CompleteAbort();
END_IF;
END_METHOD

{region 'Documentation'}
(*!
<summary>Compares independent expected values with the captured observations; called when disabled as well.</summary>
*)
{endregion}
METHOD PROTECTED ProcessAssertions
VAR_INPUT
    Enable : BOOL; //! Phase permission supplied by the owning Test Case; FALSE does not authorize progression, while observation may continue.
END_VAR
FCheckDiagnosticState(Enable := Enable,
    State := State,
    IN := TO_INT(FObserved.State),
    Expected := TO_INT(FExpected.State));

FCheckExecutionStatus(Enable := Enable,
    State := State,
    IN := TO_INT(FObserved.ExecutionStatus),
    Expected := TO_INT(FExpected.ExecutionStatus));

FCheckReady(Enable := Enable,
    State := State,
    IN := FObserved.Ready,
    Expected := FExpected.Ready);

FCheckRunning(Enable := Enable,
    State := State,
    IN := FObserved.Running,
    Expected := FExpected.Running);

FCheckCompleted(Enable := Enable,
    State := State,
    IN := FObserved.Completed,
    Expected := FExpected.Completed);

FCheckError(Enable := Enable,
    State := State,
    IN := FObserved.Error,
    Expected := FExpected.Error);

FCheckEnabled(Enable := Enable,
    State := State,
    IN := FObservedEnabled,
    Expected := FExpectedEnabled);

FCheckCommandWrites(Enable := Enable,
    State := State,
    IN := FObservedCommandWrites,
    Expected := FExpectedCommandWrites);

FCheckActualValue(Enable := Enable,
    State := State,
    IN := FObservedActualValue,
    Expected := FExpectedActualValue);

FCheckRequestedValue(Enable := Enable,
    State := State,
    IN := FObservedRequestedValue,
    Expected := FExpectedRequestedValue);

IF Enable
    AND FCheckDiagnosticState.EvaluationActive
    AND FCheckExecutionStatus.EvaluationActive
    AND FCheckReady.EvaluationActive
    AND FCheckRunning.EvaluationActive
    AND FCheckCompleted.EvaluationActive
    AND FCheckError.EvaluationActive
    AND FCheckEnabled.EvaluationActive
    AND FCheckCommandWrites.EvaluationActive
    AND FCheckActualValue.EvaluationActive
    AND FCheckRequestedValue.EvaluationActive THEN
    FCheckPerformed := TRUE;
END_IF;
END_METHOD

{region 'Documentation'}
(*!
<summary>Subjects are exercised by the test, not used as its start prerequisite.</summary>
*)
{endregion}
METHOD PROTECTED ProcessPreparations
VAR_INPUT
    // SA0033: Required hook; this scenario has no Preparation phase.
    {attribute 'analysis' := '-33'}
    Enable : BOOL; //! Phase permission supplied by the owning Test Case; FALSE does not authorize progression, while observation may continue.
END_VAR
END_METHOD

{region 'Documentation'}
(*!
<summary>Restores repeatable fixture state and resets Assertions before returning to Idle.</summary>
*)
{endregion}
METHOD PROTECTED ProcessReset
FCheckPerformed := FALSE;
FResource.Initialize(InitialValue := 2);
FSubject.Initialize(Resource := FResource);
FView := FSubject;
FCheckDiagnosticState.Reset();
FCheckExecutionStatus.Reset();
FCheckReady.Reset();
FCheckRunning.Reset();
FCheckCompleted.Reset();
FCheckError.Reset();
FCheckEnabled.Reset();
FCheckCommandWrites.Reset();
FCheckActualValue.Reset();
FCheckRequestedValue.Reset();
CompleteReset();
END_METHOD

{region 'Documentation'}
(*!
<summary>Exercises one named scenario step per call; advances only after actual Assertion evaluation.</summary>
*)
{endregion}
METHOD PROTECTED ProcessTests
VAR_INPUT
    Enable : BOOL; //! Phase permission supplied by the owning Test Case; FALSE does not authorize progression, while observation may continue.
END_VAR
IF NOT Enable THEN
    RETURN;
END_IF;

IF FCheckPerformed THEN
    FCheckPerformed := FALSE;
    IF State = CompletionWithoutReadiness THEN
        CompleteTests();
        RETURN;
    END_IF;
    NextTestState();
    IF NOT IsTestingActive THEN
        RETURN;
    END_IF;
END_IF;

CASE State OF
    FaultBeforeAction:
        FResource(Available := TRUE,
            Fault := TRUE,
            Advance := TRUE);
        FSubject(Enable := TRUE,
            TargetValue := 0);
        FExpected.State := E_State.Error;
        FExpected.ExecutionStatus := E_ExecutionStatus.Error;
        FExpected.Ready := FALSE;
        FExpected.Running := FALSE;
        FExpected.Completed := FALSE;
        FExpected.Error := TRUE;
        FExpectedEnabled := TRUE;
        FExpectedCommandWrites := 0;
        FExpectedActualValue := 2;
        FExpectedRequestedValue := 2;

    RecoveredRequest:
        FResource(Available := TRUE,
            Fault := FALSE,
            Advance := FALSE);
        FSubject(Enable := TRUE,
            TargetValue := 0);
        FExpected.State := E_State.Running;
        FExpected.ExecutionStatus := E_ExecutionStatus.Running;
        FExpected.Ready := FALSE;
        FExpected.Running := TRUE;
        FExpected.Completed := FALSE;
        FExpected.Error := FALSE;
        FExpectedEnabled := TRUE;
        FExpectedCommandWrites := 1;
        FExpectedActualValue := 2;
        FExpectedRequestedValue := 0;

    FaultDuringProgress:
        FResource(Available := TRUE,
            Fault := TRUE,
            Advance := TRUE);
        FSubject(Enable := TRUE,
            TargetValue := 0);
        FExpected.State := E_State.Error;
        FExpected.ExecutionStatus := E_ExecutionStatus.Error;
        FExpected.Ready := FALSE;
        FExpected.Running := FALSE;
        FExpected.Completed := FALSE;
        FExpected.Error := TRUE;
        FExpectedEnabled := TRUE;
        FExpectedCommandWrites := 1;
        FExpectedActualValue := 2;
        FExpectedRequestedValue := 0;

    RecoveredProgress:
        FResource(Available := TRUE,
            Fault := FALSE,
            Advance := TRUE);
        FSubject(Enable := TRUE,
            TargetValue := 0);
        FExpected.State := E_State.Running;
        FExpected.ExecutionStatus := E_ExecutionStatus.Running;
        FExpected.Ready := FALSE;
        FExpected.Running := TRUE;
        FExpected.Completed := FALSE;
        FExpected.Error := FALSE;
        FExpectedEnabled := TRUE;
        FExpectedCommandWrites := 1;
        FExpectedActualValue := 1;
        FExpectedRequestedValue := 0;

    RecoveredTarget:
        FResource(Available := TRUE,
            Fault := FALSE,
            Advance := TRUE);
        FSubject(Enable := TRUE,
            TargetValue := 0);
        FExpected.State := E_State.Completed;
        FExpected.ExecutionStatus := E_ExecutionStatus.Completed;
        FExpected.Ready := TRUE;
        FExpected.Running := FALSE;
        FExpected.Completed := TRUE;
        FExpected.Error := FALSE;
        FExpectedEnabled := TRUE;
        FExpectedCommandWrites := 1;
        FExpectedActualValue := 0;
        FExpectedRequestedValue := 0;

    FaultAfterCompletion:
        FResource(Available := TRUE,
            Fault := TRUE,
            Advance := TRUE);
        FSubject(Enable := FALSE,
            TargetValue := 0);
        FExpected.State := E_State.Error;
        FExpected.ExecutionStatus := E_ExecutionStatus.Error;
        FExpected.Ready := FALSE;
        FExpected.Running := FALSE;
        FExpected.Completed := FALSE;
        FExpected.Error := TRUE;
        FExpectedEnabled := FALSE;
        FExpectedCommandWrites := 1;
        FExpectedActualValue := 0;
        FExpectedRequestedValue := 0;

    CompletionWithoutReadiness:
        FResource(Available := FALSE,
            Fault := FALSE,
            Advance := TRUE);
        FSubject(Enable := FALSE,
            TargetValue := 0);
        FExpected.State := E_State.Completed;
        FExpected.ExecutionStatus := E_ExecutionStatus.Completed;
        FExpected.Ready := FALSE;
        FExpected.Running := FALSE;
        FExpected.Completed := TRUE;
        FExpected.Error := FALSE;
        FExpectedEnabled := FALSE;
        FExpectedCommandWrites := 1;
        FExpectedActualValue := 0;
        FExpectedRequestedValue := 0;

ELSE
    Error(Message := 'Unexpected Preparation test state.');
    RETURN;
END_CASE;

FObserved := FView.Status;
FObservedEnabled := FSubject.Enabled;

FObservedCommandWrites := FResource.CommandWriteCount;
FObservedActualValue := FResource.ActualValue;
FObservedRequestedValue := FResource.RequestedValue;
END_METHOD

END_FUNCTION_BLOCK

// ---- SelfTests/TestCases/TestSuite_Preparation/Test_PreparationMockInputs.TcPOU
{region 'Documentation'}
(*!
<summary>Checks actual PreparationMock defaults, status priority, accepted Enable and replacement of stale flags.</summary>
*)
{endregion}
FUNCTION_BLOCK Test_PreparationMockInputs EXTENDS TestCaseBase
VAR
    FSubject : PreparationMock;
    FDefaultSubject : PreparationMock;
    FObserved : ST_PreparationStatus;
    FExpected : ST_PreparationStatus;
    FObservedEnabled : BOOL;
    FExpectedEnabled : BOOL;
    FCheckPerformed : BOOL;
    FCheckDiagnosticState : AssertEqual_Int;
    FCheckExecutionStatus : AssertEqual_Int;
    FCheckReady : AssertEqual_Bool;
    FCheckRunning : AssertEqual_Bool;
    FCheckCompleted : AssertEqual_Bool;
    FCheckError : AssertEqual_Bool;
    FCheckEnabled : AssertEqual_Bool;
END_VAR
VAR CONSTANT
    DefaultInputs : E_State := E_State.Running;
    ErrorBeforeCompletion : E_State := E_State.Running + 1;
    EnabledNotReady : E_State := E_State.Running + 2;
    CompletedNotReady : E_State := E_State.Running + 3;
    ActiveWork : E_State := E_State.Running + 4;
    DisabledReady : E_State := E_State.Running + 5;
    DisabledNotReady : E_State := E_State.Running + 6;
END_VAR

SUPER^();

{region 'Documentation'}
(*!
<summary>Contributes all owned Assertion results without executing the subjects.</summary>
*)
{endregion}
METHOD PROTECTED AggregateResults
VAR_INPUT
    Aggregator : I_ResultAggregator; //! Borrowed result sink owned by the outer Test Case; add this test's checking Assertions without resetting or retaining the sink.
END_VAR
Aggregator.AddProvider(Provider := FCheckDiagnosticState);
Aggregator.AddProvider(Provider := FCheckExecutionStatus);
Aggregator.AddProvider(Provider := FCheckReady);
Aggregator.AddProvider(Provider := FCheckRunning);
Aggregator.AddProvider(Provider := FCheckCompleted);
Aggregator.AddProvider(Provider := FCheckError);
Aggregator.AddProvider(Provider := FCheckEnabled);
END_METHOD

{region 'Documentation'}
(*!
<summary>Requires valid base configuration and every owned Assertion.</summary>
*)
{endregion}
METHOD PROTECTED CheckInitialization : BOOL //! TRUE when the inherited initialization check and this concrete fixture check both accept the setup.
CheckInitialization := FALSE;
IF NOT SUPER^.CheckInitialization() THEN
    RETURN;
END_IF;
IF NOT FCheckDiagnosticState.IsInitialized
    OR NOT FCheckExecutionStatus.IsInitialized
    OR NOT FCheckReady.IsInitialized
    OR NOT FCheckRunning.IsInitialized
    OR NOT FCheckCompleted.IsInitialized
    OR NOT FCheckError.IsInitialized
    OR NOT FCheckEnabled.IsInitialized THEN
    RETURN;
END_IF;

CheckInitialization := TRUE;
END_METHOD

{region 'Documentation'}
(*!
<summary>Configures this scenario, its local subjects and named Assertions.</summary>
*)
{endregion}
METHOD PROTECTED Configure
FPreparationStateCount := 0;
FTestStateCount := 7;
FCheckPerformed := FALSE;

FCheckDiagnosticState.Initialize(Parent := THIS^,
    AssertionName := 'DiagnosticState');
FCheckExecutionStatus.Initialize(Parent := THIS^,
    AssertionName := 'ExecutionStatus');
FCheckReady.Initialize(Parent := THIS^,
    AssertionName := 'Ready');
FCheckRunning.Initialize(Parent := THIS^,
    AssertionName := 'Running');
FCheckCompleted.Initialize(Parent := THIS^,
    AssertionName := 'Completed');
FCheckError.Initialize(Parent := THIS^,
    AssertionName := 'Error');
FCheckEnabled.Initialize(Parent := THIS^,
    AssertionName := 'Enabled');
END_METHOD

{region 'Documentation'}
(*!
<summary>Ends scenario processing without issuing further resource commands.</summary>
*)
{endregion}
METHOD PROTECTED ProcessAbort
VAR_INPUT
    Enable : BOOL; //! Phase permission supplied by the owning Test Case; FALSE does not authorize progression, while observation may continue.
END_VAR
IF Enable THEN
    CompleteAbort();
END_IF;
END_METHOD

{region 'Documentation'}
(*!
<summary>Compares independent expected values with the captured observations; called when disabled as well.</summary>
*)
{endregion}
METHOD PROTECTED ProcessAssertions
VAR_INPUT
    Enable : BOOL; //! Phase permission supplied by the owning Test Case; FALSE does not authorize progression, while observation may continue.
END_VAR
FCheckDiagnosticState(Enable := Enable,
    State := State,
    IN := TO_INT(FObserved.State),
    Expected := TO_INT(FExpected.State));

FCheckExecutionStatus(Enable := Enable,
    State := State,
    IN := TO_INT(FObserved.ExecutionStatus),
    Expected := TO_INT(FExpected.ExecutionStatus));

FCheckReady(Enable := Enable,
    State := State,
    IN := FObserved.Ready,
    Expected := FExpected.Ready);

FCheckRunning(Enable := Enable,
    State := State,
    IN := FObserved.Running,
    Expected := FExpected.Running);

FCheckCompleted(Enable := Enable,
    State := State,
    IN := FObserved.Completed,
    Expected := FExpected.Completed);

FCheckError(Enable := Enable,
    State := State,
    IN := FObserved.Error,
    Expected := FExpected.Error);

FCheckEnabled(Enable := Enable,
    State := State,
    IN := FObservedEnabled,
    Expected := FExpectedEnabled);

IF Enable
    AND FCheckDiagnosticState.EvaluationActive
    AND FCheckExecutionStatus.EvaluationActive
    AND FCheckReady.EvaluationActive
    AND FCheckRunning.EvaluationActive
    AND FCheckCompleted.EvaluationActive
    AND FCheckError.EvaluationActive
    AND FCheckEnabled.EvaluationActive THEN
    FCheckPerformed := TRUE;
END_IF;
END_METHOD

{region 'Documentation'}
(*!
<summary>Subjects are exercised by the test, not used as its start prerequisite.</summary>
*)
{endregion}
METHOD PROTECTED ProcessPreparations
VAR_INPUT
    // SA0033: Required hook; this scenario has no Preparation phase.
    {attribute 'analysis' := '-33'}
    Enable : BOOL; //! Phase permission supplied by the owning Test Case; FALSE does not authorize progression, while observation may continue.
END_VAR
END_METHOD

{region 'Documentation'}
(*!
<summary>Restores repeatable fixture state and resets Assertions before returning to Idle.</summary>
*)
{endregion}
METHOD PROTECTED ProcessReset
FCheckPerformed := FALSE;
FCheckDiagnosticState.Reset();
FCheckExecutionStatus.Reset();
FCheckReady.Reset();
FCheckRunning.Reset();
FCheckCompleted.Reset();
FCheckError.Reset();
FCheckEnabled.Reset();
CompleteReset();
END_METHOD

{region 'Documentation'}
(*!
<summary>Exercises one named scenario step per call; advances only after actual Assertion evaluation.</summary>
*)
{endregion}
METHOD PROTECTED ProcessTests
VAR_INPUT
    Enable : BOOL; //! Phase permission supplied by the owning Test Case; FALSE does not authorize progression, while observation may continue.
END_VAR
IF NOT Enable THEN
    RETURN;
END_IF;

IF FCheckPerformed THEN
    FCheckPerformed := FALSE;
    IF State = DisabledNotReady THEN
        CompleteTests();
        RETURN;
    END_IF;
    NextTestState();
    IF NOT IsTestingActive THEN
        RETURN;
    END_IF;
END_IF;

CASE State OF
    DefaultInputs:
        FDefaultSubject(Enable := FALSE);
        FObserved := FDefaultSubject.Status;
        FObservedEnabled := FDefaultSubject.Enabled;
        FExpected.State := E_State.Completed;
        FExpected.ExecutionStatus := E_ExecutionStatus.Completed;
        FExpected.Ready := TRUE;
        FExpected.Running := FALSE;
        FExpected.Completed := TRUE;
        FExpected.Error := FALSE;
        FExpectedEnabled := FALSE;

    ErrorBeforeCompletion:
        FSubject(Enable := TRUE,
            Ready := TRUE,
            Completed := TRUE,
            Error := TRUE);
        FObserved := FSubject.Status;
        FObservedEnabled := FSubject.Enabled;
        FExpected.State := E_State.Error;
        FExpected.ExecutionStatus := E_ExecutionStatus.Error;
        FExpected.Ready := TRUE;
        FExpected.Running := FALSE;
        FExpected.Completed := FALSE;
        FExpected.Error := TRUE;
        FExpectedEnabled := TRUE;

    EnabledNotReady:
        FSubject(Enable := TRUE,
            Ready := FALSE,
            Completed := FALSE,
            Error := FALSE);
        FObserved := FSubject.Status;
        FObservedEnabled := FSubject.Enabled;
        FExpected.State := E_State.Idle;
        FExpected.ExecutionStatus := E_ExecutionStatus.NotReady;
        FExpected.Ready := FALSE;
        FExpected.Running := FALSE;
        FExpected.Completed := FALSE;
        FExpected.Error := FALSE;
        FExpectedEnabled := TRUE;

    CompletedNotReady:
        FSubject(Enable := TRUE,
            Ready := FALSE,
            Completed := TRUE,
            Error := FALSE);
        FObserved := FSubject.Status;
        FObservedEnabled := FSubject.Enabled;
        FExpected.State := E_State.Completed;
        FExpected.ExecutionStatus := E_ExecutionStatus.Completed;
        FExpected.Ready := FALSE;
        FExpected.Running := FALSE;
        FExpected.Completed := TRUE;
        FExpected.Error := FALSE;
        FExpectedEnabled := TRUE;

    ActiveWork:
        FSubject(Enable := TRUE,
            Ready := TRUE,
            Completed := FALSE,
            Error := FALSE);
        FObserved := FSubject.Status;
        FObservedEnabled := FSubject.Enabled;
        FExpected.State := E_State.Running;
        FExpected.ExecutionStatus := E_ExecutionStatus.Running;
        FExpected.Ready := FALSE;
        FExpected.Running := TRUE;
        FExpected.Completed := FALSE;
        FExpected.Error := FALSE;
        FExpectedEnabled := TRUE;

    DisabledReady:
        FSubject(Enable := FALSE,
            Ready := TRUE,
            Completed := FALSE,
            Error := FALSE);
        FObserved := FSubject.Status;
        FObservedEnabled := FSubject.Enabled;
        FExpected.State := E_State.Idle;
        FExpected.ExecutionStatus := E_ExecutionStatus.Idle;
        FExpected.Ready := TRUE;
        FExpected.Running := FALSE;
        FExpected.Completed := FALSE;
        FExpected.Error := FALSE;
        FExpectedEnabled := FALSE;

    DisabledNotReady:
        FSubject(Enable := FALSE,
            Ready := FALSE,
            Completed := FALSE,
            Error := FALSE);
        FObserved := FSubject.Status;
        FObservedEnabled := FSubject.Enabled;
        FExpected.State := E_State.Idle;
        FExpected.ExecutionStatus := E_ExecutionStatus.NotReady;
        FExpected.Ready := FALSE;
        FExpected.Running := FALSE;
        FExpected.Completed := FALSE;
        FExpected.Error := FALSE;
        FExpectedEnabled := FALSE;

ELSE
    Error(Message := 'Unexpected Preparation test state.');
    RETURN;
END_CASE;
END_METHOD

END_FUNCTION_BLOCK

// ---- Framework/Preparation/POU/PreparationMock.TcPOU
{region 'Documentation'}
(*!
<summary>Controllable Preparation double without resource actions or automatic
progression.</summary>
<description>
On each call, Error takes priority over Completed, then Enabled AND Ready selects Running;
otherwise Ready selects Idle or NotReady. Completion is observed independently of Enable and is not
latched.

Defaults Ready=TRUE, Completed=TRUE and Error=FALSE report a reached target after the first
call. Before that call, Status retains its uninitialized defaults.
</description>
*)
{endregion}
FUNCTION_BLOCK PreparationMock EXTENDS PreparationBase
VAR_INPUT
    Ready : BOOL := TRUE; //! Simulated resource readiness; the reported status suppresses Ready while Running. Does not mean target reached.
    Completed : BOOL := TRUE; //! Preparation target is currently reached; observation is not latched.
    Error : BOOL := FALSE; //! Preparation cannot continue meaningfully; reported as an error observation.
END_VAR

SUPER^();

{region 'Documentation'}
(*!
<summary>Reflect inputs on every call; Error overrides Completed, then active work; otherwise Ready
selects Idle or NotReady.</summary>
*)
{endregion}
METHOD PROTECTED Prepare
IF Error THEN
    UpdateStatus(State := E_State.Error,
        ExecutionStatus := E_ExecutionStatus.Error,
        Ready := Ready);
    RETURN;
END_IF;

IF Completed THEN
    UpdateStatus(State := E_State.Completed,
        ExecutionStatus := E_ExecutionStatus.Completed,
        Ready := Ready);
    RETURN;
END_IF;

IF Enabled AND Ready THEN
    UpdateStatus(State := E_State.Running,
        ExecutionStatus := E_ExecutionStatus.Running,
        Ready := FALSE);
    RETURN;
END_IF;

IF NOT Ready THEN
    UpdateStatus(State := E_State.Idle,
        ExecutionStatus := E_ExecutionStatus.NotReady,
        Ready := FALSE);
    RETURN;
END_IF;

UpdateStatus(State := E_State.Idle,
    ExecutionStatus := E_ExecutionStatus.Idle,
    Ready := Ready);
END_METHOD

END_FUNCTION_BLOCK

// ---- SelfTests/TestSuites/TestSuite_TestCaseLifecycle.TcPOU
{region 'Documentation'}
(*!
<summary>Verifies the real Test Case lifecycle through isolated subjects and serial checking Test Cases.</summary>
*)
{endregion}
FUNCTION_BLOCK TestSuite_TestCaseLifecycle EXTENDS TestSuiteBase
VAR
    FInitialization : Test_LifecycleInitialization;
    FWithoutPreparation : Test_LifecycleWithoutPreparation;
    FSinglePreparation : Test_LifecycleSinglePreparation;
    FMultipleStates : Test_LifecycleMultipleStates;
    FAlreadyPrepared : Test_LifecycleAlreadyPrepared;
    FFailedResult : Test_LifecycleFailedResult;
    FAbort : Test_LifecycleAbort;
    FAbortError : Test_LifecycleAbortError;
    FAbortTimeout : Test_LifecycleAbortTimeout;
    FExecutionTimeout : Test_LifecycleExecutionTimeout;
    FPreparationError : Test_LifecyclePreparationError;
    FPreparationTimeout : Test_LifecyclePreparationTimeout;
    FResetError : Test_LifecycleResetError;
    FResetTimeout : Test_LifecycleResetTimeout;
    FResetDuringExecution : Test_LifecycleResetDuringExecution;
    FFailedToError : Test_LifecycleFailedToError;
    FInvalidTestAdvance : Test_LifecycleInvalidTestAdvance;
    FInvalidPreparationTransition : Test_LifecycleInvalidPreparationTransition;
    FRepeatAfterPassed : Test_LifecycleRepeatAfterPassed;
    FRepeatAfterFailed : Test_LifecycleRepeatAfterFailed;
    FRepeatAfterError : Test_LifecycleRepeatAfterError;
    FRepeatAfterAbort : Test_LifecycleRepeatAfterAbort;
    FTestCases : ARRAY[1..TestCaseCapacity] OF I_TestCase;
END_VAR
VAR CONSTANT
    TestCaseCapacity : UINT := 22;
END_VAR

SUPER^();

{region 'Documentation'}
(*!
<summary>Binds subject identity before outer initialization and registers deterministic serial order.</summary>
*)
{endregion}
METHOD PROTECTED Configure
VAR_IN_OUT
    // SA0167: Borrowed builder; VAR_IN_OUT creates no temporary instance.
    {attribute 'analysis' := '-167'}
    Builder : TestSuiteConfigurationBuilder; //! Borrowed owner configuration builder used only during this Configure call; register this owner's concrete children.
END_VAR
VAR
    TestConfig : ST_TestCaseConfig;
END_VAR
Builder.Initialize(Mode := E_OrchestrationMode.Serial,
    TestCases := FTestCases);

FInitialization.BindSubjectParent(Parent := THIS^);
FInitialization.Initialize(Parent := THIS^,
    TestName := 'Initialization',
    Config := TestConfig);
Builder.Register(TestCase := FInitialization);

FWithoutPreparation.BindSubjectParent(Parent := THIS^);
FWithoutPreparation.Initialize(Parent := THIS^,
    TestName := 'WithoutPreparation',
    Config := TestConfig);
Builder.Register(TestCase := FWithoutPreparation);

FSinglePreparation.BindSubjectParent(Parent := THIS^);
FSinglePreparation.Initialize(Parent := THIS^,
    TestName := 'SinglePreparation',
    Config := TestConfig);
Builder.Register(TestCase := FSinglePreparation);

FMultipleStates.BindSubjectParent(Parent := THIS^);
FMultipleStates.Initialize(Parent := THIS^,
    TestName := 'MultipleStates',
    Config := TestConfig);
Builder.Register(TestCase := FMultipleStates);

FAlreadyPrepared.BindSubjectParent(Parent := THIS^);
FAlreadyPrepared.Initialize(Parent := THIS^,
    TestName := 'AlreadyPrepared',
    Config := TestConfig);
Builder.Register(TestCase := FAlreadyPrepared);

FFailedResult.BindSubjectParent(Parent := THIS^);
FFailedResult.Initialize(Parent := THIS^,
    TestName := 'FailedResult',
    Config := TestConfig);
Builder.Register(TestCase := FFailedResult);

FAbort.BindSubjectParent(Parent := THIS^);
FAbort.Initialize(Parent := THIS^,
    TestName := 'Abort',
    Config := TestConfig);
Builder.Register(TestCase := FAbort);

FAbortError.BindSubjectParent(Parent := THIS^);
FAbortError.Initialize(Parent := THIS^,
    TestName := 'AbortError',
    Config := TestConfig);
Builder.Register(TestCase := FAbortError);

FAbortTimeout.BindSubjectParent(Parent := THIS^);
FAbortTimeout.Initialize(Parent := THIS^,
    TestName := 'AbortTimeout',
    Config := TestConfig);
Builder.Register(TestCase := FAbortTimeout);

FExecutionTimeout.BindSubjectParent(Parent := THIS^);
FExecutionTimeout.Initialize(Parent := THIS^,
    TestName := 'ExecutionTimeout',
    Config := TestConfig);
Builder.Register(TestCase := FExecutionTimeout);

FPreparationError.BindSubjectParent(Parent := THIS^);
FPreparationError.Initialize(Parent := THIS^,
    TestName := 'PreparationError',
    Config := TestConfig);
Builder.Register(TestCase := FPreparationError);

FPreparationTimeout.BindSubjectParent(Parent := THIS^);
FPreparationTimeout.Initialize(Parent := THIS^,
    TestName := 'PreparationTimeout',
    Config := TestConfig);
Builder.Register(TestCase := FPreparationTimeout);

FResetError.BindSubjectParent(Parent := THIS^);
FResetError.Initialize(Parent := THIS^,
    TestName := 'ResetError',
    Config := TestConfig);
Builder.Register(TestCase := FResetError);

FResetTimeout.BindSubjectParent(Parent := THIS^);
FResetTimeout.Initialize(Parent := THIS^,
    TestName := 'ResetTimeout',
    Config := TestConfig);
Builder.Register(TestCase := FResetTimeout);

FResetDuringExecution.BindSubjectParent(Parent := THIS^);
FResetDuringExecution.Initialize(Parent := THIS^,
    TestName := 'ResetDuringExecution',
    Config := TestConfig);
Builder.Register(TestCase := FResetDuringExecution);

FFailedToError.BindSubjectParent(Parent := THIS^);
FFailedToError.Initialize(Parent := THIS^,
    TestName := 'FailedToError',
    Config := TestConfig);
Builder.Register(TestCase := FFailedToError);

FInvalidTestAdvance.BindSubjectParent(Parent := THIS^);
FInvalidTestAdvance.Initialize(Parent := THIS^,
    TestName := 'InvalidTestAdvance',
    Config := TestConfig);
Builder.Register(TestCase := FInvalidTestAdvance);

FInvalidPreparationTransition.BindSubjectParent(Parent := THIS^);
FInvalidPreparationTransition.Initialize(Parent := THIS^,
    TestName := 'InvalidPreparationTransition',
    Config := TestConfig);
Builder.Register(TestCase := FInvalidPreparationTransition);

FRepeatAfterPassed.BindSubjectParent(Parent := THIS^);
FRepeatAfterPassed.Initialize(Parent := THIS^,
    TestName := 'RepeatAfterPassed',
    Config := TestConfig);
Builder.Register(TestCase := FRepeatAfterPassed);

FRepeatAfterFailed.BindSubjectParent(Parent := THIS^);
FRepeatAfterFailed.Initialize(Parent := THIS^,
    TestName := 'RepeatAfterFailed',
    Config := TestConfig);
Builder.Register(TestCase := FRepeatAfterFailed);

FRepeatAfterError.BindSubjectParent(Parent := THIS^);
FRepeatAfterError.Initialize(Parent := THIS^,
    TestName := 'RepeatAfterError',
    Config := TestConfig);
Builder.Register(TestCase := FRepeatAfterError);

FRepeatAfterAbort.BindSubjectParent(Parent := THIS^);
FRepeatAfterAbort.Initialize(Parent := THIS^,
    TestName := 'RepeatAfterAbort',
    Config := TestConfig);
Builder.Register(TestCase := FRepeatAfterAbort);
END_METHOD

{region 'Documentation'}
(*!
<summary>Resolves the same array that Configure registered.</summary>
*)
{endregion}
METHOD PUBLIC GetTestCase : I_TestCase //! Typed child interface at the original array index; zero when no entry is available.
VAR_INPUT
    Index : DINT; //! Original occupied child-array index, rather than an ordinal position.
END_VAR
GetTestCase := 0;
IF (ChildCount = 0) OR (Index < ChildArrayLowerBound)
    OR (DINT_TO_LINT(Index) >= DINT_TO_LINT(ChildArrayLowerBound) + UINT_TO_LINT(ChildCount)) THEN
    RETURN;
END_IF;
GetTestCase := FTestCases[Index];
END_METHOD

{region 'Documentation'}
(*!
<summary>Calls each owned checking Test Case once per initialized Suite cycle.</summary>
*)
{endregion}
METHOD PROTECTED ProcessTestCases
FInitialization();
FWithoutPreparation();
FSinglePreparation();
FMultipleStates();
FAlreadyPrepared();
FFailedResult();
FAbort();
FAbortError();
FAbortTimeout();
FExecutionTimeout();
FPreparationError();
FPreparationTimeout();
FResetError();
FResetTimeout();
FResetDuringExecution();
FFailedToError();
FInvalidTestAdvance();
FInvalidPreparationTransition();
FRepeatAfterPassed();
FRepeatAfterFailed();
FRepeatAfterError();
FRepeatAfterAbort();
END_METHOD

END_FUNCTION_BLOCK

// ---- SelfTests/TestCases/TestSuite_TestCaseLifecycle/Test_LifecycleInitialization.TcPOU
{region 'Documentation'}
(*!
<summary>Checks identity/configuration rejection and passivity before the first lifecycle Reset.</summary>
<description>
Each Test state is one initialization attempt with an independent local event capture.
BeginAttempt varies exactly one configuration condition. Identity errors must stop before
Configure; setup errors must reach Configure while the subject is still Uninitialized.
Two later subject calls verify that rejected objects remain passive and do not repeat
initialization diagnostics. Start/Abort are submitted only before the first call. A valid
initialized subject emits their two Trigger events but must still wait for its parent's
Reset; the following call must not repeat either requests or initialization diagnostics.
The checking Assertions retain failures across all attempts and publish normally.
</description>
*)
{endregion}
FUNCTION_BLOCK Test_LifecycleInitialization EXTENDS TestCaseBase
VAR
    FSubjectParent : I_TestSuite;
    FSubject : TestCaseInitializationProbe;
    FCapture : EventBuffer;
    FEvents : ARRAY[1..CaptureLength] OF ST_Event;
    FCaptureFifo : ST_FifoStatus;
    FCaptureStatus : ST_EventBufferStatus;
    FFixtureValid : BOOL;
    FAttempt : INT := 1;
    FAttemptStarted : BOOL;
    FCheckPerformed : BOOL;
    FPassiveCallCount : UINT;
    FExpectedInitialized : BOOL;
    FExpectedConfigured : BOOL;
    FInitializationMatches : BOOL;
    FConfigureOrderMatches : BOOL;
    FDiagnosticMatches : BOOL;
    FPassiveStateMatches : BOOL;
    FHookCallsMatch : BOOL;
    FEventsUnchanged : BOOL;
    FSequenceAfterInitialize : UDINT;
    FCheckInitialization : AssertTrue;
    FCheckConfigureOrder : AssertTrue;
    FCheckPassiveState : AssertTrue;
    FCheckHookDispatch : AssertTrue;
    FCheckDiagnostic : AssertTrue;
    FCheckNoRepeatedEvents : AssertTrue;
    FCheckCaptureIntegrity : AssertTrue;
END_VAR
VAR CONSTANT
    CaptureLength : UINT := 32;
    PassiveCallCount : UINT := 2;
    RequestTriggerCount : UDINT := 2;
    MissingParent : INT := 1;
    InvalidSegment : INT := 2;
    OverlengthName : INT := 3;
    UnconfiguredPreparations : INT := 4;
    UnconfiguredTests : INT := 5;
    NegativePreparationCount : INT := 6;
    ExcessPreparationCount : INT := 7;
    NoTestStates : INT := 8;
    ExcessTestCount : INT := 9;
    ZeroExecutionTimeout : INT := 10;
    ZeroPreparationTimeout : INT := 11;
    ZeroResetTimeout : INT := 12;
    ZeroAbortTimeout : INT := 13;
    ConcreteRejection : INT := 14;
    ValidConfiguration : INT := 15;
    AttemptCount : INT := 15;
END_VAR

SUPER^();

{region 'Documentation'}
(*!
<summary>Supplies the seven checking results; expected subject errors are not outer errors.</summary>
*)
{endregion}
METHOD PROTECTED AggregateResults
VAR_INPUT
    Aggregator : I_ResultAggregator; //! Borrowed result sink owned by the outer Test Case; add this test's checking Assertions without resetting or retaining the sink.
END_VAR
Aggregator.AddProvider(Provider := FCheckInitialization);
Aggregator.AddProvider(Provider := FCheckConfigureOrder);
Aggregator.AddProvider(Provider := FCheckPassiveState);
Aggregator.AddProvider(Provider := FCheckHookDispatch);
Aggregator.AddProvider(Provider := FCheckDiagnostic);
Aggregator.AddProvider(Provider := FCheckNoRepeatedEvents);
Aggregator.AddProvider(Provider := FCheckCaptureIntegrity);
END_METHOD

{region 'Documentation'}
(*!
<summary>Varies one input; records immediate Initialize evidence before any cyclic subject call.</summary>
*)
{endregion}
METHOD PRIVATE BeginAttempt
VAR
    Config : ST_TestCaseConfig;
    Parent : I_TestSuite;
    TestName : STRING(GVL_Constants.NameLength);
    PreparationCount : INT;
    TestCount : INT := 1;
    Initialized : BOOL;
    Index : UINT;
END_VAR
FFixtureValid := FCapture.Initialize(Buffer := FEvents,
    FifoControl := FCaptureFifo,
    Status := FCaptureStatus);
IF NOT FFixtureValid THEN
    Error(Message := 'Initialization test capture could not be initialized.');
    RETURN;
END_IF;

Parent := FSubjectParent;
TestName := 'Subject';
CASE FAttempt OF
    MissingParent:
        Parent := 0;
    InvalidSegment:
        TestName := 'Invalid.Subject';
    OverlengthName:
        FOR Index := 1 TO GVL_Constants.NameLength DO
            TestName := CONCAT(TestName, 'x');
        END_FOR;
    UnconfiguredPreparations:
        PreparationCount := -1;
    UnconfiguredTests:
        TestCount := -1;
    NegativePreparationCount:
        PreparationCount := -2;
    ExcessPreparationCount:
        PreparationCount := E_State.Running - E_State.Preparing + 1;
    NoTestStates:
        TestCount := 0;
    ExcessTestCount:
        TestCount := E_State.Completing - E_State.Running + 1;
    ZeroExecutionTimeout:
        Config.Timeout := T#0s;
    ZeroPreparationTimeout:
        Config.PreparationTimeout := T#0s;
    ZeroResetTimeout:
        Config.ResetTimeout := T#0s;
    ZeroAbortTimeout:
        Config.AbortTimeout := T#0s;
END_CASE;

FExpectedInitialized := FAttempt = ValidConfiguration;
FExpectedConfigured := FAttempt >= UnconfiguredPreparations;
FSubject.BeginScenario(RejectConfiguration := FAttempt = ConcreteRejection);
FSubject.Bind(Publisher := FCapture,
    PreparationCount := PreparationCount,
    TestCount := TestCount);
Initialized := FSubject.Initialize(Parent := Parent,
    TestName := TestName,
    Config := Config);
FInitializationMatches := (Initialized = FExpectedInitialized)
    AND (FSubject.IsInitialized = FExpectedInitialized);
FConfigureOrderMatches := FSubject.WasConfigured() = FExpectedConfigured;
IF FExpectedConfigured THEN
    FConfigureOrderMatches := FConfigureOrderMatches AND FSubject.WasConfigurationContextValid();
END_IF;

FSequenceAfterInitialize := FCaptureStatus.SequenceId;
IF FExpectedInitialized THEN
    FDiagnosticMatches := FSequenceAfterInitialize = 0;
ELSE
    FDiagnosticMatches := (FSequenceAfterInitialize = 1)
        AND (FEvents[1].Severity = E_EventSeverity.Error)
        AND (FEvents[1].State = E_State.Uninitialized);
    IF FAttempt = MissingParent THEN
        FDiagnosticMatches := FDiagnosticMatches AND (FEvents[1].Name = TestName);
    ELSE
        FDiagnosticMatches := FDiagnosticMatches AND (FEvents[1].Name = FSubject.Name);
    END_IF;
END_IF;
FPassiveStateMatches := TRUE;
FHookCallsMatch := TRUE;
FEventsUnchanged := TRUE;
FPassiveCallCount := 0;
FAttemptStarted := TRUE;
END_METHOD

{region 'Documentation'}
(*!
<summary>Supplies identity only; the containing Suite never executes the isolated subject.</summary>
*)
{endregion}
METHOD PUBLIC BindSubjectParent
VAR_INPUT
    Parent : I_TestSuite; //! Borrowed identity parent retained for isolated subject initialization; keep the Suite alive through subject use.
END_VAR
FSubjectParent := Parent;
END_METHOD

{region 'Documentation'}
(*!
<summary>Initializes the outer Assertions; subject initialization is the test action, not fixture setup.</summary>
*)
{endregion}
METHOD PROTECTED Configure
FPreparationStateCount := 0;
FTestStateCount := AttemptCount;
FCheckInitialization.Initialize(Parent := THIS^,
    AssertionName := 'Initialization');
FCheckConfigureOrder.Initialize(Parent := THIS^,
    AssertionName := 'ConfigureOrder');
FCheckPassiveState.Initialize(Parent := THIS^,
    AssertionName := 'PassiveState');
FCheckHookDispatch.Initialize(Parent := THIS^,
    AssertionName := 'HookDispatch');
FCheckDiagnostic.Initialize(Parent := THIS^,
    AssertionName := 'Diagnostic');
FCheckNoRepeatedEvents.Initialize(Parent := THIS^,
    AssertionName := 'NoRepeatedEvents');
FCheckCaptureIntegrity.Initialize(Parent := THIS^,
    AssertionName := 'CaptureIntegrity');
END_METHOD

{region 'Documentation'}
(*!
<summary>The test owns no asynchronous resource action.</summary>
*)
{endregion}
METHOD PROTECTED ProcessAbort
VAR_INPUT
    Enable : BOOL; //! Phase permission supplied by the owning Test Case; FALSE does not authorize progression, while observation may continue.
END_VAR
IF Enable THEN
    CompleteAbort();
END_IF;
END_METHOD

{region 'Documentation'}
(*!
<summary>Latches each attempt&#x27;s independent checks in the outer Assertions.</summary>
*)
{endregion}
METHOD PROTECTED ProcessAssertions
VAR_INPUT
    Enable : BOOL; //! Phase permission supplied by the owning Test Case; FALSE does not authorize progression, while observation may continue.
END_VAR
VAR
    Evaluate : BOOL;
END_VAR
Evaluate := Enable AND (FPassiveCallCount >= PassiveCallCount);
FCheckInitialization(Enable := Evaluate,
    State := FState,
    IN := FInitializationMatches);
FCheckConfigureOrder(Enable := Evaluate,
    State := FState,
    IN := FConfigureOrderMatches);
FCheckPassiveState(Enable := Evaluate,
    State := FState,
    IN := FPassiveStateMatches);
FCheckHookDispatch(Enable := Evaluate,
    State := FState,
    IN := FHookCallsMatch);
FCheckDiagnostic(Enable := Evaluate,
    State := FState,
    IN := FDiagnosticMatches);
FCheckNoRepeatedEvents(Enable := Evaluate,
    State := FState,
    IN := FEventsUnchanged);
FCheckCaptureIntegrity(Enable := Evaluate,
    State := FState,
    IN := NOT FSubject.TraceOverflow AND (FCaptureStatus.LostEventCount = 0));
IF Evaluate THEN
    FCheckPerformed := TRUE;
END_IF;
END_METHOD

{region 'Documentation'}
(*!
<summary>No preparation phase is required.</summary>
*)
{endregion}
METHOD PROTECTED ProcessPreparations
VAR_INPUT
    {attribute 'analysis' := '-33'}
    Enable : BOOL; //! Phase permission supplied by the owning Test Case; FALSE does not authorize progression, while observation may continue.
END_VAR
END_METHOD

{region 'Documentation'}
(*!
<summary>Restarts the attempts and resets checking Assertions without initializing the subject.</summary>
*)
{endregion}
METHOD PROTECTED ProcessReset
FAttempt := 1;
FAttemptStarted := FALSE;
FCheckPerformed := FALSE;
FPassiveCallCount := 0;
FCheckInitialization.Reset();
FCheckConfigureOrder.Reset();
FCheckPassiveState.Reset();
FCheckHookDispatch.Reset();
FCheckDiagnostic.Reset();
FCheckNoRepeatedEvents.Reset();
FCheckCaptureIntegrity.Reset();
CompleteReset();
END_METHOD

{region 'Documentation'}
(*!
<summary>Calls the subject once per active PLC cycle; checks span two calls before advancing.</summary>
*)
{endregion}
METHOD PROTECTED ProcessTests
VAR_INPUT
    Enable : BOOL; //! Phase permission supplied by the owning Test Case; FALSE does not authorize progression, while observation may continue.
END_VAR
VAR
    HookIndex : UINT;
    Hook : ST_LifecycleHook;
END_VAR
IF NOT Enable THEN
    RETURN;
END_IF;
IF FCheckPerformed THEN
    IF FAttempt = AttemptCount THEN
        CompleteTests();
        RETURN;
    END_IF;
    FAttempt := FAttempt + 1;
    FAttemptStarted := FALSE;
    FCheckPerformed := FALSE;
    NextTestState();
END_IF;
IF NOT FAttemptStarted THEN
    BeginAttempt();
    IF NOT FFixtureValid THEN
        RETURN;
    END_IF;
END_IF;

// Start/Abort cannot bypass the required parent Reset, whether setup succeeded or failed.
IF FPassiveCallCount = 0 THEN
    FSubject.RequestStart();
    FSubject.RequestAbort();
END_IF;
FSubject();
FPassiveStateMatches := FPassiveStateMatches
    AND (FSubject.State = E_State.Uninitialized)
    AND NOT FSubject.IsReady
    AND (FSubject.Result = E_Result.NotEvaluated);
IF FExpectedInitialized THEN
    FHookCallsMatch := FHookCallsMatch AND (FSubject.HookCount = 5);
    FOR HookIndex := 1 TO FSubject.HookCount DO
        Hook := FSubject.GetHook(Index := HookIndex);
        IF Hook.Hook <> E_LifecycleHook.Aggregate THEN
            FHookCallsMatch := FHookCallsMatch AND NOT Hook.Enabled;
        END_IF;
    END_FOR;
ELSE
    FHookCallsMatch := FHookCallsMatch AND (FSubject.HookCount = 0);
END_IF;
IF FExpectedInitialized THEN
    FEventsUnchanged := FEventsUnchanged
        AND (FCaptureStatus.SequenceId = FSequenceAfterInitialize + RequestTriggerCount)
        AND (FEvents[1].EventType = E_EventType.Trigger)
        AND (FEvents[1].Name = FSubject.Name)
        AND (FEvents[1].State = E_State.Uninitialized)
        AND (FEvents[1].Message = 'Abort trigger.')
        AND (FEvents[2].EventType = E_EventType.Trigger)
        AND (FEvents[2].Name = FSubject.Name)
        AND (FEvents[2].State = E_State.Uninitialized)
        AND (FEvents[2].Message = 'Start trigger.');
ELSE
    FEventsUnchanged := FEventsUnchanged AND (FCaptureStatus.SequenceId = FSequenceAfterInitialize);
END_IF;
FPassiveCallCount := FPassiveCallCount + 1;
END_METHOD

END_FUNCTION_BLOCK

// ---- SelfTests/TestCases/TestSuite_TestCaseLifecycle/Helper/TestCaseInitializationProbe.TcPOU
{region 'Documentation'}
(*!
<summary>Observes initialization ordering without replacing the production lifecycle.</summary>
<description>
BeginScenario clears only this adapter's observations. Configure records the state in which
the production Initialize calls it. The optional rejection exercises a concrete owner's
additional CheckInitialization failure after the inherited checks have passed.
</description>
*)
{endregion}
FUNCTION_BLOCK TestCaseInitializationProbe EXTENDS TestCaseLifecycleProbe
VAR
    FConfigurationObserved : BOOL;
    FConfigurationContextValid : BOOL;
    FRejectConfiguration : BOOL;
END_VAR

SUPER^();

{region 'Documentation'}
(*!
<summary>Clears observations before one explicit initialization attempt.</summary>
*)
{endregion}
METHOD PUBLIC BeginScenario
VAR_INPUT
    RejectConfiguration : BOOL := FALSE; //! TRUE makes the concrete initialization check report Error and reject configuration.
END_VAR
FConfigurationObserved := FALSE;
FConfigurationContextValid := FALSE;
FRejectConfiguration := RejectConfiguration;
END_METHOD

{region 'Documentation'}
(*!
<summary>Rejects a concrete setup only after the inherited checks succeeded.</summary>
*)
{endregion}
METHOD PROTECTED CheckInitialization : BOOL //! TRUE when the inherited initialization check and this concrete fixture check both accept the setup.
CheckInitialization := FALSE;
IF NOT SUPER^.CheckInitialization() THEN
    RETURN;
END_IF;
IF FRejectConfiguration THEN
    EventPublisher.PublishEvent(Event := CreateFrameworkEvent(Name := Name,
        ResourceName := FResourceName,
        State := State,
        Severity := E_EventSeverity.Error,
        Message := 'Concrete test setup rejected.'));
    RETURN;
END_IF;
CheckInitialization := TRUE;
END_METHOD

{region 'Documentation'}
(*!
<summary>Observes entry, then uses the existing concrete hook implementation.</summary>
*)
{endregion}
METHOD PROTECTED Configure
FConfigurationObserved := TRUE;
FConfigurationContextValid := (State = E_State.Uninitialized) AND NOT IsInitialized AND (Name <> '');
SUPER^.Configure();
END_METHOD

{region 'Documentation'}
(*!
<summary>Configure must run with the new identity, Uninitialized state and initialization not yet accepted.</summary>
*)
{endregion}
METHOD PUBLIC WasConfigurationContextValid : BOOL //! Recorded TRUE when Configure observed the expected new identity and pre-acceptance initialization context.
WasConfigurationContextValid := FConfigurationContextValid;
END_METHOD

{region 'Documentation'}
(*!
<summary>Reports whether Configure was reached in this initialization attempt.</summary>
*)
{endregion}
METHOD PUBLIC WasConfigured : BOOL //! TRUE when Configure was reached during the current scenario.
WasConfigured := FConfigurationObserved;
END_METHOD

END_FUNCTION_BLOCK

// ---- SelfTests/TestCases/TestSuite_TestCaseLifecycle/Helper/TestCaseLifecycleProbe.TcPOU
{region 'Documentation'}
(*!
<summary>
Provides controllable application hooks around the unchanged TestCaseBase lifecycle.
</summary>

<description>

Controlled behavior

Inputs emulate concrete application decisions inside the Process* overrides.
The overrides call the real base APIs for errors and phase completion;
they do not replace the Sequencer or assign its state directly.
Two real Assertions provide child results: Condition is controlled,
while ReferenceCondition always receives TRUE.

Per-call trace

Each override records method, state and Enable before performing its action.
A transition inside one hook is visible when the following hook records its entry.
The FB call clears the previous trace before invoking SUPER^().
The fixed trace buffer belongs to this probe, not to the event stream.

Binding and evaluation

Bind supplies the isolated publisher and phase counts before Initialize.
The outer TestCaseLifecycleTestBase drives this object and judges its observations;
the subject's own result is test data, not the outer selftest verdict.
</description>
*)
{endregion}
FUNCTION_BLOCK TestCaseLifecycleProbe EXTENDS TestCaseBase
VAR_INPUT
    Ready : BOOL := TRUE; //! Scenario readiness release, combined with inherited startability.
    ResetCompleted : BOOL := TRUE; //! TRUE permits the Reset hook to report completion.
    PreparationTargetReached : BOOL := FALSE; //! Scripted preparation target condition.
    AdvancePreparation : BOOL := FALSE; //! TRUE permits the preparation hook to advance its state.
    FinishPreparations : BOOL := FALSE; //! TRUE permits the preparation hook to complete its phase.
    AdvanceTest : BOOL := FALSE; //! TRUE permits the test hook to advance its state.
    FinishTests : BOOL := FALSE; //! TRUE permits the test hook to complete its phase.
    AssertionCondition : BOOL := TRUE; //! Condition supplied to the controlled Assertion.
    AbortCompleted : BOOL := TRUE; //! TRUE permits the Abort hook to report completion.
    ResetError : BOOL := FALSE; //! TRUE injects a technical Error from the Reset hook.
    TestError : BOOL := FALSE; //! TRUE injects a technical Error from the test hook.
    AbortError : BOOL := FALSE; //! TRUE injects a technical Error from the Abort hook.
    PreparationError : BOOL := FALSE; //! TRUE injects a technical Error from the preparation hook.
END_VAR
VAR
    FConfiguredPreparationCount : INT;
    FConfiguredTestCount : INT := 1;
    FAssertion : AssertTrue;
    FReferenceAssertion : AssertTrue;
    FHooks : ARRAY[1..HookCapacity] OF ST_LifecycleHook;
    FHookCount : UINT;
    FTraceOverflow : BOOL;
END_VAR
VAR CONSTANT
    HookCapacity : UINT := 6;
END_VAR

// Keep only this call's observations; SUPER^ invokes the instrumented overrides below.
FHookCount := 0;
FTraceOverflow := FALSE;
SUPER^();

{region 'Documentation'}
(*!
<summary>Contributes both real child results; the inherited base owns interpretation and counters.</summary>
*)
{endregion}
METHOD PROTECTED AggregateResults
VAR_INPUT
    Aggregator : I_ResultAggregator; //! Borrowed result sink owned by the outer Test Case; add this test's checking Assertions without resetting or retaining the sink.
END_VAR
RecordHook(Hook := E_LifecycleHook.Aggregate,
    Enabled := TRUE);
Aggregator.AddProvider(Provider := FAssertion);
Aggregator.AddProvider(Provider := FReferenceAssertion);
END_METHOD

{region 'Documentation'}
(*!
<summary>Selects publisher and scenario shape before calling the inherited Initialize.</summary>
*)
{endregion}
METHOD PUBLIC Bind
VAR_INPUT
    Publisher : I_EventPublisher; //! Nonzero isolated event publisher retained before subject initialization; keep it alive through all subject use.
    PreparationCount : INT; //! Preparation-state count supplied to the next concrete Configure call.
    TestCount : INT; //! Test-state count supplied to the next concrete Configure call.
END_VAR
FEventPublisher := Publisher;
FConfiguredPreparationCount := PreparationCount;
FConfiguredTestCount := TestCount;
FAssertion.BindPublisher(Publisher := Publisher);
FReferenceAssertion.BindPublisher(Publisher := Publisher);
END_METHOD

{region 'Documentation'}
(*!
<summary>Keeps the base validation and rejects an unusable owned Assertion.</summary>
*)
{endregion}
METHOD PROTECTED CheckInitialization : BOOL //! TRUE when the inherited initialization check and this concrete fixture check both accept the setup.
CheckInitialization := SUPER^.CheckInitialization()
    AND FAssertion.IsInitialized AND FReferenceAssertion.IsInitialized;
END_METHOD

{region 'Documentation'}
(*!
<summary>Initializes the two real Assertions and configures the requested phase counts.</summary>
*)
{endregion}
METHOD PROTECTED Configure
FPreparationStateCount := FConfiguredPreparationCount;
FTestStateCount := FConfiguredTestCount;
FHookCount := 0;
FTraceOverflow := FALSE;
FAssertion.Initialize(Parent := THIS^,
    AssertionName := 'Condition');
FReferenceAssertion.Initialize(Parent := THIS^,
    AssertionName := 'ReferenceCondition');
END_METHOD

{region 'Documentation'}
(*!
<summary>Returns the recorded entry; an invalid index returns the empty observation.</summary>
*)
{endregion}
METHOD PUBLIC GetHook : ST_LifecycleHook //! Recorded hook entry at Index; an empty entry when Index is outside 1..HookCount.
VAR_INPUT
    Index : UINT; //! One-based hook-entry index within 1..HookCount; other indices return an empty entry.
END_VAR
VAR
    EmptyHook : ST_LifecycleHook;
END_VAR
GetHook := EmptyHook;
IF (Index < 1) OR (Index > FHookCount) THEN
    RETURN;
END_IF;

GetHook := FHooks[Index];
END_METHOD

